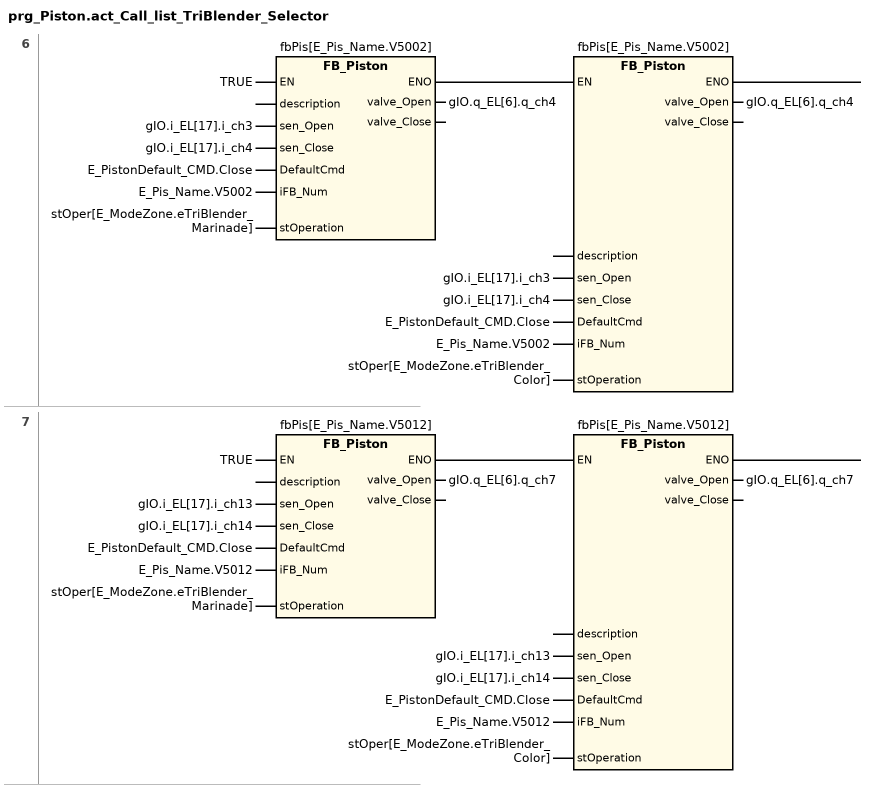
// NETWORK 6
fbPis[E_Pis_Name.V5002](
    sen_Open := gIO.i_EL[17].i_ch3,
    sen_Close := gIO.i_EL[17].i_ch4,
    DefaultCmd := E_PistonDefault_CMD.Close,
    iFB_Num := E_Pis_Name.V5002,
    stOperation := stOper[E_ModeZone.eTriBlender_Marinade],
    valve_Open => gIO.q_EL[6].q_ch4); // FB_Piston
fbPis[E_Pis_Name.V5002](
    sen_Open := gIO.i_EL[17].i_ch3,
    sen_Close := gIO.i_EL[17].i_ch4,
    DefaultCmd := E_PistonDefault_CMD.Close,
    iFB_Num := E_Pis_Name.V5002,
    stOperation := stOper[E_ModeZone.eTriBlender_Color],
    valve_Open => gIO.q_EL[6].q_ch4); // FB_Piston

// NETWORK 7
fbPis[E_Pis_Name.V5012](
    sen_Open := gIO.i_EL[17].i_ch13,
    sen_Close := gIO.i_EL[17].i_ch14,
    DefaultCmd := E_PistonDefault_CMD.Close,
    iFB_Num := E_Pis_Name.V5012,
    stOperation := stOper[E_ModeZone.eTriBlender_Marinade],
    valve_Open => gIO.q_EL[6].q_ch7); // FB_Piston
fbPis[E_Pis_Name.V5012](
    sen_Open := gIO.i_EL[17].i_ch13,
    sen_Close := gIO.i_EL[17].i_ch14,
    DefaultCmd := E_PistonDefault_CMD.Close,
    iFB_Num := E_Pis_Name.V5012,
    stOperation := stOper[E_ModeZone.eTriBlender_Color],
    valve_Open => gIO.q_EL[6].q_ch7); // FB_Piston
END_ACTION

ACTION act_Call_list_Water:
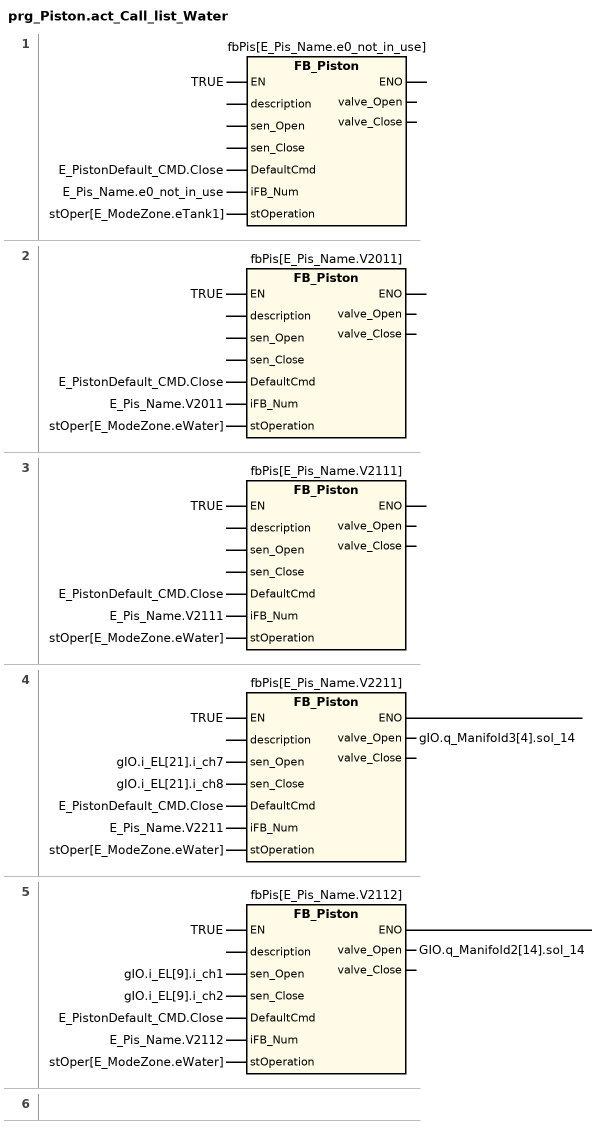
// NETWORK 1
fbPis[E_Pis_Name.e0_not_in_use](
    DefaultCmd := E_PistonDefault_CMD.Close,
    iFB_Num := E_Pis_Name.e0_not_in_use,
    stOperation := stOper[E_ModeZone.eTank1]); // FB_Piston

// NETWORK 2
fbPis[E_Pis_Name.V2011](
    DefaultCmd := E_PistonDefault_CMD.Close,
    iFB_Num := E_Pis_Name.V2011,
    stOperation := stOper[E_ModeZone.eWater]); // FB_Piston

// NETWORK 3
fbPis[E_Pis_Name.V2111](
    DefaultCmd := E_PistonDefault_CMD.Close,
    iFB_Num := E_Pis_Name.V2111,
    stOperation := stOper[E_ModeZone.eWater]); // FB_Piston

// NETWORK 4
fbPis[E_Pis_Name.V2211](
    sen_Open := gIO.i_EL[21].i_ch7,
    sen_Close := gIO.i_EL[21].i_ch8,
    DefaultCmd := E_PistonDefault_CMD.Close,
    iFB_Num := E_Pis_Name.V2211,
    stOperation := stOper[E_ModeZone.eWater],
    valve_Open => gIO.q_Manifold3[4].sol_14); // FB_Piston

// NETWORK 5
fbPis[E_Pis_Name.V2112](
    sen_Open := gIO.i_EL[9].i_ch1,
    sen_Close := gIO.i_EL[9].i_ch2,
    DefaultCmd := E_PistonDefault_CMD.Close,
    iFB_Num := E_Pis_Name.V2112,
    stOperation := stOper[E_ModeZone.eWater],
    valve_Open => GIO.q_Manifold2[14].sol_14); // FB_Piston

// NETWORK 6
END_ACTION

ACTION act_InterLock:
(*
IF TRUE 
AND stPis[E_Pis_Name.cheesy_cut].st_Deafult
AND stPis[E_Pis_Name.cheesy_down].st_Deafult
AND stPis[E_Pis_Name.cheesy_gripper].st_Deafult
AND stPis[E_Pis_Name.cheesy_turn].st_Deafult

AND stPis[E_Pis_Name.crown_down].st_Deafult
AND stPis[E_Pis_Name.crown_gripper].st_Deafult
AND stPis[E_Pis_Name.crown_press].st_Deafult
AND stPis[E_Pis_Name.crown_push].st_Deafult

AND stPis[E_Pis_Name.crust_down].st_Deafult
AND stPis[E_Pis_Name.crust_hold].st_Deafult
AND stPis[E_Pis_Name.crust_push].st_Deafult
AND stPis[E_Pis_Name.crust_roll].st_Deafult

AND stPis[E_Pis_Name.spikes_rotate_4].st_Deafult
AND stPis[E_Pis_Name.spikes_updown_4].st_Deafult

AND stPis[E_Pis_Name.door_4_2].st_Deafult

AND stPis[E_Pis_Name.trolley_down].st_Deafult

THEN;
	stPis[E_Pis_Name.trolley_move].b_InterLock:=TRUE;
ELSE;
	stPis[E_Pis_Name.trolley_move].b_InterLock:=FALSE;
END_IF
*)
END_ACTION

METHOD m_Disable_All : BOOL
VAR_INPUT
END_VAR

VAR
	i: INT;
END_VAR
FOR i:=1 TO E_Pis_Name.last DO;
	stPis[i].b_Enable:=FALSE;
END_FOR
END_METHOD

METHOD m_Enable_All : BOOL
VAR_INPUT
END_VAR

VAR
	i: INT;
END_VAR
FOR i:=1 TO E_Pis_Name.last DO;
	stPis[i].b_Enable:=TRUE;
END_FOR
END_METHOD

METHOD m_Get_Next_N : BOOL
VAR_IN_OUT
	iSel: INT;
END_VAR

VAR
	i: INT;
END_VAR

IF iSel> 1 THEN;
	FOR i:=iSel-1 TO 1 BY -1 DO
		IF stPis[i].b_Exist THEN;
			iSel:=i;
			RETURN;
		END_IF		
	END_FOR
END_IF
END_METHOD

METHOD m_Get_Next_P : BOOL
VAR_IN_OUT
	iSel: INT;
END_VAR

VAR
	i: INT;
END_VAR
//IF iSel< C_MAX_Pistons THEN;
//IF iSel< C_MAX_Pistons_Exist THEN;
IF iSel< E_Pis_Name.last THEN;
	FOR i:=iSel+1 TO E_Pis_Name.last BY 1 DO
		IF stPis[i].b_Exist THEN;
			iSel:=i;
			RETURN;
		END_IF		
	END_FOR
END_IF
END_METHOD

END_PROGRAM

// ---- 00 Library/01 Piston/FB_Piston.TcPOU
FUNCTION_BLOCK FB_Piston
VAR_INPUT
	description		: STRING;		(* Piston description*)	
	sen_Open		: BOOL;
	sen_Close		: BOOL;
	
	DefaultCmd		: E_PistonDefault_CMD:=E_PistonDefault_CMD.Close;

	iFB_Num			: E_Pis_Name;

END_VAR
VAR_OUTPUT
	valve_Open		: BOOL;
	valve_Close		: BOOL;	
END_VAR
VAR_IN_OUT
	stOperation		: ST_OperationButtons;	
END_VAR
VAR
	stPis			:	REFERENCE TO ST_Piston;
	stPis_UpLow		:	REFERENCE TO ST_Piston_U_L;
	state: E_Piston_State;
	state_Close,state_Open: (Ready, CheckState, ValveUpdate, Busy, Delay, Done, Error);

	//sen_Open_Exist	: REFERENCE TO BOOL :=FALSE;
	//sen_Close_Exist	: REFERENCE TO BOOL :=FALSE;
	
	ton_SensorCheck	: TON;
	ton_MinTime		: TON;
	ton_MaxTime		: TON;
	ton_SensorDelay	: TON;

	// Timing 
	t_minOpen		: TIME 	:=T#300MS;	(* minimum time to open piston*)
	t_minClose		: TIME	:=T#300MS;	(* minimum time to close piston*)
	t_maxOpen		: TIME 	:=T#3S;		(* Maximum time to open piston, will initiate an error*)
	t_maxClose		: TIME	:=T#3S;		(* Maximum time to open piston, will initiate an error*)
	t_DelayOpen		: TIME 	:=T#0S;		(* Delay time to getting "st_Open", will count after minimum time and sensors detection done*)
	t_DelayClose	: TIME	:=T#0S;		(* Delay time to getting "st_Close", will count after minimum time and sensors detection done*)	
	
	rt_Close		: R_TRIG;
	rt_Open			: R_TRIG;
	rt_OpenMan		: R_TRIG;
	rt_CloseMan		: R_TRIG;
	rt_DefaultPos	: R_TRIG;
	rt_ResumeMaster	: R_TRIG;
	b_memo_OpenFDBKExist	: BOOL;
	b_memo_CloseFDBKExist	: BOOL;
	Call_FTrig_ReqUp	: F_TRIG;
	Call_FTrig_ReqLow	: F_TRIG;
	
	bErrorMemo: BOOL;
		
	ton_Req_Close_timeout: TON;
	ton_Req_Open_timeout: TON;
	ton_Req_Default_timeout: TON;
	rt_StateSafe: R_TRIG;
	ft_StateSafe: F_TRIG;
END_VAR

IF iFB_Num <> E_Pis_Name.e0_not_in_use THEN;
	
END_IF

act_Get_Reference();




act_State_Machine();
act_StateDeafult();
//act_MemFdbkExist();

stPis_UpLow.bError:=stPis.b_Error;
stPis_UpLow.iFB_Num:=iFB_Num;
	
IF iFB_Num = E_Pis_Name.e0_not_in_use THEN;
	//stPis.st_Deafult:=TRUE;
END_IF


rt_StateSafe(CLK:=stOperation.bStateSafe_mode);
ft_StateSafe(CLK:=stOperation.bStateSafe_mode);

IF __ISVALIDREF(stPis) THEN;
	IF ft_StateSafe.Q
	AND NOT stPis.st_Deafult
	THEN;
		//stPis.req_DefaultPos:=TRUE;
		//stPis.req_Close:=FALSE;
		//stPis.req_Open:=FALSE;	
	END_IF
	
	IF rt_StateSafe.Q THEN;
		
		IF NOT stPis.st_Deafult THEN;
			//stPis.req_DefaultPos:=TRUE;
		END_IF	
		stPis.b_Resume:=TRUE;
		//stPis.b_Reset:=TRUE;	
	END_IF	
END_IF

ACTION act_Close:



CASE state_Close OF
	Ready:;
		IF stPis.req_CloseMan THEN;
			stPis.req_CloseMan:=FALSE;
			// Do manual case code
			stPis.req_Close:=TRUE;
		END_IF		
		IF stPis.req_Close THEN;
			stPis.req_Open:=FALSE;
			stPis.req_OpenMan:=FALSE;	
			stPis.req_DefaultPos:=FALSE;			
			state_Close:=CheckState;
		END_IF
		
	CheckState:;
		IF stPis.st_Close THEN;
			stPis.st_Open:=FALSE;
			state_Close:=Done;
		ELSE;
			stPis.st_Close:=FALSE;
			stPis.st_Open:=FALSE;
			state_Close:=ValveUpdate;
		END_IF
		
	ValveUpdate:;
		valve_Open:=FALSE;
		valve_Close:=TRUE;
		ton_SensorCheck(IN:=FALSE);
		ton_MinTime(IN:=FALSE);
		ton_MinTime(IN:=TRUE);
		ton_MaxTime(IN:=FALSE);
		ton_MaxTime(IN:=TRUE);
		ton_SensorDelay(IN:=FALSE);
		
		stPis.t_LastClose:=T#0S;
		state_Close:=Busy;
		
	Busy:;
		ton_MinTime(PT:=t_minClose);
		ton_MaxTime(PT:=t_maxClose, IN:=TRUE);
		ton_SensorDelay(PT:=t_DelayClose,IN:=m_PistonSensorCheck());	
		IF 	ton_MinTime.Q 		
		AND ton_SensorDelay.IN THEN;
			ton_MaxTime(IN:=FALSE);
			IF ton_SensorDelay.Q THEN;
				stPis.t_LastClose:=ton_MaxTime.ET;			
				state_Close:=Done;				
			END_IF
		ELSE;
			IF ton_MaxTime.Q THEN;
				//Error to print
				state_Close:=Error;
			END_IF			
		END_IF
	
	Done:;
		stPis.st_Close:=TRUE;
		IF stPis.st_Close THEN;
			state_Close:=Ready;
			stPis.req_Close:=FALSE;
		END_IF	
		
	Error:;
		//Wating to operator reset & resume 
		stPis.b_Error:=TRUE;	
		m_Error();
		IF stPis.b_Resume THEN;
			state_Close:=ValveUpdate;
			//stPis.b_Resume:=FALSE;	
			//stPis.b_Error:=FALSE;
			//bErrorMemo:=FALSE;
		END_IF
		
END_CASE
END_ACTION

ACTION act_Get_Reference:
stPis REF= g_Piston.stPis[iFB_Num];
stPis_UpLow REF= g_Piston.stPis_U_L[iFB_Num];
//stPis.description:=description;
stPis.b_Exist:=TRUE;
stPis.sName:=TO_STRING(iFB_Num);
stPis.iPisNum:=iFB_Num;
arPisName[iFB_Num].Num:=iFB_Num;
arPisName[iFB_Num].Description:=stPis.sName;

stPis.sen_Close REF= sen_Close;
stPis.sen_Close_Exist REF= stPisSetting[iFB_Num].sen_Close_Exist;
//stPis.sen_Close_Exist REF= sen_Close_Exist;
stPis.sen_Open REF= sen_Open;
stPis.sen_Open_Exist REF= stPisSetting[iFB_Num].sen_Open_Exist;
//stPis.sen_Open_Exist REF= sen_Open_Exist;

stPis.valve_Close REF= valve_Close;
stPis.valve_Open REF= valve_Open;

stPis.t_maxClose REF= stPisSetting[iFB_Num].t_maxClose;
stPis.t_maxOpen REF= stPisSetting[iFB_Num].t_maxOpen;
stPis.t_minClose REF= stPisSetting[iFB_Num].t_minClose;
stPis.t_minOpen REF= stPisSetting[iFB_Num].t_minOpen;
stPis.t_DelayClose REF= stPisSetting[iFB_Num].t_DelayClose;
stPis.t_DelayOpen REF= stPisSetting[iFB_Num].t_DelayOpen;
t_maxClose:=fun_Real_SecondsToTime(in_Time:=stPis.t_maxClose);
t_maxOpen:=fun_Real_SecondsToTime(in_Time:=stPis.t_maxOpen);
t_minClose:=fun_Real_SecondsToTime(in_Time:=stPis.t_minClose);
t_minOpen:=fun_Real_SecondsToTime(in_Time:=stPis.t_minOpen);
t_DelayClose:=fun_Real_SecondsToTime(in_Time:=stPis.t_DelayClose);
t_DelayOpen:=fun_Real_SecondsToTime(in_Time:=stPis.t_DelayOpen);

stPis.DefaultCmd REF= DefaultCmd;

IF stPis.b_Error THEN;
	stOperation.bSetPause:=TRUE;
END_IF
(*
IF stPis.b_Error 
AND stDevErr_H.eErrorActive=E_Error_Active_Module.noError 
THEN;
	stDevErr_H.sObjectName:=CONCAT('pis.No:',INT_TO_STRING(stPis.iPisNum));
	stDevErr_H.sObjectName:=CONCAT(stDevErr_H.sObjectName,'- ');
	stDevErr_H.sObjectName:=CONCAT(stDevErr_H.sObjectName,TO_STRING(iFB_Num));
	stDevErr_H.eErrorActive:=E_Error_Active_Module.Piston;
	stDevErr_H.iObjectID:=iFB_Num;
END_IF

rt_ResumeMaster(CLK:=stDevErr_H.bMasterResume);
IF rt_ResumeMaster.Q THEN;
	stPis.b_Resume:=TRUE;
END_IF
*)
END_ACTION

ACTION act_MemFdbkExist:
IF stPis.valve_Close AND stPis_UpLow.exist THEN
	//Fetching signals
	IF TRUE THEN
		Call_FTrig_ReqUp(CLK:=stPis_UpLow.req_Upper , Q=> );
	ELSE
		Call_FTrig_ReqUp(CLK:=stPis_UpLow.st_Upper , Q=> );
	END_IF
	
	Call_FTrig_ReqLow(CLK:=stPis_UpLow.st_Lower , Q=> );
	
	//setting memmory
	IF stPis_UpLow.req_Lower AND stPis.sen_Close_Exist THEN
		b_memo_CloseFDBKExist:=stPis.sen_Close_Exist;
		stPis.sen_Close_Exist:=FALSE;
	ELSIF stPis_UpLow.req_Lower AND b_memo_CloseFDBKExist THEN
		stPis.sen_Close_Exist:=FALSE;
	END_IF
	
	IF stPis_UpLow.req_Upper AND stPis.sen_Open_Exist THEN
		b_memo_OpenFDBKExist:=stPis.sen_Open_Exist;
		stPis.sen_Open_Exist:=FALSE;
	ELSIF stPis_UpLow.req_Upper AND b_memo_OpenFDBKExist THEN
		stPis.sen_Open_Exist:=FALSE;
	END_IF
	//resseting memmory
	IF Call_FTrig_ReqUp.Q AND b_memo_OpenFDBKExist THEN
		stPis.sen_Open_Exist:=b_memo_OpenFDBKExist;
		b_memo_OpenFDBKExist:=FALSE;
	END_IF
	
	IF Call_FTrig_ReqLow.Q AND b_memo_CloseFDBKExist THEN
		stPis.sen_Close_Exist:=b_memo_CloseFDBKExist;
		b_memo_CloseFDBKExist:=FALSE;
	END_IF
ELSE
	IF stPis_UpLow.exist THEN
		b_memo_CloseFDBKExist:=FALSE;
		b_memo_OpenFDBKExist:=FALSE;
		stPis_UpLow.req_Lower:=FALSE;
		stPis_UpLow.st_Lower:=FALSE;
	ELSE
		;
	END_IF
	
END_IF

IF stPis.req_Open AND NOT stPis_UpLow.exist  THEN
	IF stPis.sen_Close_Exist THEN
		b_memo_CloseFDBKExist:=TRUE;
		stPis.sen_Close_Exist:=FALSE;
	END_IF
	
	IF stPis.sen_Open_Exist THEN
		b_memo_OpenFDBKExist:=TRUE;
		stPis.sen_Open_Exist:=FALSE;
	END_IF
ELSIF stPis.req_Close AND NOT stPis_UpLow.exist THEN
	IF b_memo_CloseFDBKExist THEN
		stPis.sen_Close_Exist:=TRUE;
		b_memo_CloseFDBKExist:=FALSE;
	END_IF
	
	IF b_memo_OpenFDBKExist THEN
		stPis.sen_Open_Exist:=TRUE;
		b_memo_OpenFDBKExist:=FALSE;
	END_IF
	
END_IF
END_ACTION

ACTION act_New_CMD:
IF stPis.b_Enable AND stPis.b_InterLock THEN;
	
	rt_Close(CLK:=stPis.req_Close AND NOT ton_Req_Close_timeout.Q);
	rt_Open(CLK:=stPis.req_Open AND NOT ton_Req_Open_timeout.Q);
	rt_CloseMan(CLK:=stPis.req_CloseMan);
	rt_OpenMan(CLK:=stPis.req_OpenMan);
	rt_DefaultPos(CLK:=stPis.req_DefaultPos AND NOT ton_Req_Default_timeout.Q);
	
	ton_Req_Close_timeout(PT:=T#0.1S);	
	IF (stPis.req_Close OR stPis.req_CloseMan)
	AND state_Close=Ready
	AND NOT ton_Req_Close_timeout.Q
	THEN;
		ton_Req_Close_timeout.IN:=TRUE;
	ELSE;
		ton_Req_Close_timeout.IN:=FALSE;
	END_IF

	ton_Req_Open_timeout(PT:=T#0.1S);	
	IF (stPis.req_Open OR stPis.req_OpenMan)
	AND state_Open=Ready
	AND NOT ton_Req_Open_timeout.Q
	THEN;
		ton_Req_Open_timeout.IN:=TRUE;
	ELSE;
		ton_Req_Open_timeout.IN:=FALSE;
	END_IF

	ton_Req_Default_timeout(PT:=T#0.1S);	
	IF (stPis.req_DefaultPos OR stPis.req_DefaultPos)
	AND state_Open=Ready
	AND NOT ton_Req_Default_timeout.Q
	THEN;
		ton_Req_Default_timeout.IN:=TRUE;
	ELSE;
		ton_Req_Default_timeout.IN:=FALSE;
	END_IF
	
	IF rt_Close.Q OR rt_CloseMan.Q THEN; 
		state:=E_Piston_State.Busy_Close; 
		stPis.req_Open:=FALSE;
		stPis.req_OpenMan:=FALSE;	
		stPis.req_DefaultPos:=FALSE;	
	END_IF
	IF rt_Open.Q OR rt_OpenMan.Q THEN; 
		state:=E_Piston_State.Busy_Open; 
		stPis.req_Close:=FALSE;
		stPis.req_CloseMan:=FALSE;
		stPis.req_DefaultPos:=FALSE;	
	END_IF
	IF rt_DefaultPos.Q THEN; 
		state:=E_Piston_State.Init; 
	END_IF
	
	(*IF rt_CloseMan.Q THEN; 
		state:=E_Piston_State.Busy_Close;
	END_IF
	IF rt_OpenMan.Q THEN; 
		state:=E_Piston_State.Busy_Open; 
	END_IF
*)
	
	IF rt_Close.Q 
	OR rt_Open.Q
	OR rt_CloseMan.Q
	OR rt_OpenMan.Q
	OR rt_DefaultPos.Q
	THEN;
		stPis.b_Error:=FALSE;
		bErrorMemo:=FALSE;
	END_IF
	
	stPis.b_DeactivateMan:=FALSE;
ELSE;
	stPis.b_DeactivateMan:=TRUE;
END_IF
END_ACTION

ACTION act_Open:



CASE state_Open OF
	Ready:;
		IF stPis.req_OpenMan THEN;
			stPis.req_OpenMan:=FALSE;
			// Do manual case code
			stPis.req_Open:=TRUE;
		END_IF		
		IF stPis.req_Open THEN;
			stPis.req_Close:=FALSE;
			stPis.req_CloseMan:=FALSE;
			stPis.req_DefaultPos:=FALSE;		
			state_Open:=CheckState;
		END_IF
		
	CheckState:;
		IF stPis.st_Open THEN;
			stPis.st_Close:=FALSE;
			state_Open:=Done;
		ELSE;
			stPis.st_Close:=FALSE;
			stPis.st_Open:=FALSE;
			state_Open:=ValveUpdate;
		END_IF
		
	ValveUpdate:;
		valve_Open:=TRUE;
		valve_Close:=FALSE;
		ton_SensorCheck(IN:=FALSE);
		ton_MinTime(IN:=FALSE);
		ton_MinTime(IN:=TRUE);
		ton_MaxTime(IN:=FALSE);
		ton_MaxTime(IN:=TRUE);	
		ton_SensorDelay(IN:=FALSE);
		
		stPis.t_LastOpen:=T#0S;	
		state_Open:=Busy;
		
	Busy:;
		ton_MinTime(PT:=t_minOpen);
		ton_MaxTime(PT:=t_maxOpen);
		ton_SensorDelay(PT:=t_DelayOpen,IN:=m_PistonSensorCheck());	
		IF 	ton_MinTime.Q 
		AND m_PistonSensorCheck()	THEN;
			ton_MaxTime(IN:=FALSE);
			IF ton_SensorDelay.Q THEN;
				stPis.t_LastOpen:=ton_MaxTime.ET;			
				state_Open:=Done;				
			END_IF
		ELSE;
			IF ton_MaxTime.Q THEN;
				//Error to print
				state_Open:=Error;
				;
			END_IF				
		END_IF
	
	Done:;
		stPis.st_Open:=TRUE;	
		IF stPis.st_Open THEN;
			state_Open:=Ready;
			stPis.req_Open:=FALSE;
		END_IF	
		
	Error:;
		//Wating to operator reset & resume 
		stPis.b_Error:=TRUE;
		m_Error();
		IF stPis.b_Resume THEN;
			state_Open:=ValveUpdate;
			//stPis.b_Resume:=FALSE;
			//stPis.b_Error:=FALSE;
			//bErrorMemo:=FALSE;
		END_IF
		
END_CASE
END_ACTION

ACTION act_State_Machine:
IF stPis.b_Resume THEN;
	stPis.b_Error:=FALSE;
	bErrorMemo:=FALSE;		
END_IF

act_New_CMD();
CASE state OF
	E_Piston_State.Init:;
			ton_SensorCheck(IN:=FALSE);
			
	
			stPis.st_Close:=FALSE;
			stPis.st_Open:=FALSE;
			
			stPis.b_Error:=FALSE;
			stPis.b_Reset:=FALSE;
			stPis.b_Resume:=FALSE;
			
			stPis.req_Close:=FALSE;
			stPis.req_CloseMan:=FALSE;	
			stPis.req_Open:=FALSE;
			stPis.req_OpenMan:=FALSE;
			stPis.req_DefaultPos:=FALSE;
			
			state_Close:=Ready;
			state_Open:=Ready;
			
			//check default configuration
			IF stPis.b_Enable AND stPis.b_InterLock THEN;				
				CASE DefaultCmd OF
					E_PistonDefault_CMD.Close:;
						state:=E_Piston_State.Busy_Close;
						stPis.req_Close:=TRUE;
					E_PistonDefault_CMD.Open:;
						state:=E_Piston_State.Busy_Open;
						stPis.req_Open:=TRUE;
					E_PistonDefault_CMD.Sensors:;
					E_PistonDefault_CMD.SensorsClose:;
					E_PistonDefault_CMD.SensorsOpen:;
					
				END_CASE
			END_IF
	
	E_Piston_State.Close:;
		IF m_PistonSensorCheck() AND NOT stPis.b_Error THEN;
			stPis.st_Close:=TRUE;
			stPis.st_Open:=FALSE;
			ton_SensorCheck(IN:=FALSE);
		ELSE;
			ton_SensorCheck(IN:=TRUE);
			IF ton_SensorCheck.Q THEN;
				stPis.st_Close:=FALSE;
				stPis.st_Open:=FALSE;				
				stPis.b_Error:=TRUE;
				m_Error();		
			END_IF			
		END_IF
				
	E_Piston_State.Open:;
		IF m_PistonSensorCheck() AND NOT stPis.b_Error THEN;
			stPis.st_Close:=FALSE;
			stPis.st_Open:=TRUE;
			ton_SensorCheck(IN:=FALSE);
		ELSE;			
			ton_SensorCheck(IN:=TRUE);
			IF ton_SensorCheck.Q THEN;
				stPis.st_Close:=FALSE;
				stPis.st_Open:=FALSE;				
				stPis.b_Error:=TRUE;
				m_Error();
			END_IF
		END_IF
	
	E_Piston_State.Busy_Close:;
		ton_SensorCheck(IN:=FALSE);
		act_Close();		
		state_Open:=Ready;		
		IF stPis.st_Close AND NOT stPis.req_Close THEN;
			state:=E_Piston_State.Close;
		END_IF

	E_Piston_State.Busy_Open:;
		ton_SensorCheck(IN:=FALSE);
		act_Open();
		state_Close:=Ready;
		IF stPis.st_Open AND NOT stPis.req_Open THEN;
			state:=E_Piston_State.Open;
		END_IF
END_CASE			

ton_SensorCheck(PT:=T#4S);//PT:=T#0.5S

IF ton_SensorCheck.Q THEN;
	stPis.b_Error:=TRUE;		
END_IF
stPis.b_Resume:=FALSE;
END_ACTION

ACTION act_StateDeafult:
CASE DefaultCmd	OF
	E_PistonDefault_CMD.Close:;
		stPis.st_Deafult:=stPis.st_Close;
	E_PistonDefault_CMD.Open:;
		stPis.st_Deafult:=stPis.st_Open;
END_CASE
END_ACTION

METHOD PUBLIC m_CheckByRecipe : BOOL
VAR_INPUT
	stPis: ST_Piston;
	req: E_Piston_Recipe_State;	
END_VAR
m_CheckByRecipe:=FALSE;
IF stPis.iPisNum <> E_Pis_Name.e0_not_in_use THEN
	CASE req OF
		E_Piston_Recipe_State.NoChanges:;
			m_CheckByRecipe:=TRUE;
		E_Piston_Recipe_State.Act:;
			IF (stPis.DefaultCmd=E_PistonDefault_CMD.Close AND stPis.st_Open) 
			OR (stPis.DefaultCmd=E_PistonDefault_CMD.Open AND stPis.st_Close)
			THEN;
				m_CheckByRecipe:=TRUE;
			END_IF
		E_Piston_Recipe_State.Release:;
			IF (stPis.DefaultCmd=E_PistonDefault_CMD.Close AND stPis.st_Close) 
			OR (stPis.DefaultCmd=E_PistonDefault_CMD.Open AND stPis.st_Open)
			THEN;
				m_CheckByRecipe:=TRUE;
			END_IF	
	END_CASE
ELSE;
	m_CheckByRecipe:=TRUE;
END_IF
END_METHOD

METHOD m_Error : BOOL
VAR_INPUT
END_VAR
VAR
	sActErrorID_AA: STRING;
	sActErrorID: STRING;
	Mess: INT;
	cFound: INT;
	iFound: INT;
	i: INT;
	bWarning: BOOL;

END_VAR
(*
IF SFCError OR bWarning THEN

	IF  SFCErrorStep='WaitSenOpen' THEN
		stPis.eErrNum:=1;
	ELSIF SFCErrorStep='WaitSenNotClose' THEN
		stPis.eErrNum:=2;
	ELSIF SFCErrorStep='WaitSenClose' THEN
		stPis.eErrNum:=3;
	ELSIF SFCErrorStep='WaitSenNotOpen' THEN
		stPis.eErrNum:=4;
	ELSIF SFCErrorStep='No Status' THEN
		stPis.eErrNum:=5;
	ELSIF SFCErrorStep='No Valve Operation' THEN
		stPis.eErrNum:=6;
	ELSIF SFCErrorStep='Not synchronized with cycle command' THEN //SensorsChecking
		stPis.eErrNum:=7;
	ELSIF SFCErrorStep='SensorsChecking' THEN
		stPis.eErrNum:=8;		
	ELSIF bWarning THEN;	// act_Ready
		//stPis.eErrNum:=21; 	// '2AAx021',	'Warning',	', Manual command rejected in semi/auto mode',	(**)
	ELSE
		stPis.eErrNum:=9;
	END_IF
	Last_SFCErrorStep:=SFCErrorStep;
	
ELSE
		stPis.eErrNum:=0;
END_IF
*)
// Temp solution
IF stPis.b_Error THEN;
	stPis.eErrNum:=1;
END_IF

IF stPis.eErrNum<>0 AND NOT bErrorMemo AND stPis.iPisNum<>0 THEN

	IF stPis.iPisNum<10 THEN
		sActErrorID:=CONCAT('20',INT_TO_STRING(stPis.iPisNum));
	ELSE
		sActErrorID:=CONCAT('2',INT_TO_STRING(stPis.iPisNum));
	END_IF
	
	IF stPis.eErrNum<10 THEN
		sActErrorID:=CONCAT(sActErrorID,'x00');
		sActErrorID:=CONCAT(sActErrorID,INT_TO_STRING(stPis.eErrNum));
	ELSE
		sActErrorID:=CONCAT(sActErrorID,'x0');
		sActErrorID:=CONCAT(sActErrorID,INT_TO_STRING(stPis.eErrNum));		
	END_IF

	FOR Mess:=100 TO 2 BY -1 DO
		Buffer_Act_Message[Mess].sDateTime:=Buffer_Act_Message[Mess-1].sDateTime;
		Buffer_Act_Message[Mess].sErrID:=Buffer_Act_Message[Mess-1].sErrID;
		Buffer_Act_Message[Mess].sLevel:=Buffer_Act_Message[Mess-1].sLevel;
		Buffer_Act_Message[Mess].sModuleDescription:=Buffer_Act_Message[Mess-1].sModuleDescription;
		Buffer_Act_Message[Mess].sErrorMessage:=Buffer_Act_Message[Mess-1].sErrorMessage;
	END_FOR
		Buffer_Act_Message[1].sDateTime:=sRealTime;
		Buffer_Act_Message[1].sErrID:=sActErrorID;
		Buffer_Act_Message[1].sLevel:='Error';
		//Buffer_Act_Message[1].sModuleDescription:='Pneumatic valve';
		Buffer_Act_Message[1].sModuleDescription:=stOperation.sModeZone;

		(*888888888888888888888888888888888888888888*)
		IF stPis.eErrNum<10 THEN
			sActErrorID_AA:=CONCAT('2AAx00',INT_TO_STRING(stPis.eErrNum));
		ELSE
			sActErrorID_AA:=CONCAT('2AAx0',INT_TO_STRING(stPis.eErrNum));			
		END_IF
		cFound:=0;
		FOR i:=1 TO C_Max_ErrorList DO
			IF ar_ErrorList[i,eErrID]=sActErrorID_AA THEN
				iFound:=i;
				ar_ErrorActive[iFound]:=TRUE;
				cFound:=cFound+1;
			END_IF
		END_FOR

		Buffer_Act_Message[1].sErrorMessage:=CONCAT( 'Piston Num ', INT_TO_STRING(stPis.iPisNum));
		Buffer_Act_Message[1].sErrorMessage:=CONCAT( Buffer_Act_Message[1].sErrorMessage, ', ');
		//Buffer_Act_Message[1].sErrorMessage:=CONCAT( Buffer_Act_Message[1].sErrorMessage, arPisDescription[stPis.iPisNum]);
		Buffer_Act_Message[1].sErrorMessage:=CONCAT( Buffer_Act_Message[1].sErrorMessage, stPis.sName);
		Buffer_Act_Message[1].sErrorMessage:=CONCAT( Buffer_Act_Message[1].sErrorMessage, ': ');

		IF cFound=1 THEN;
			Buffer_Act_Message[1].sErrorMessage:=CONCAT( Buffer_Act_Message[1].sErrorMessage, ar_ErrorList[iFound,eErrMeassage]);	(*	Error from the List	*)
			Buffer_Act_Message[1].sLevel:= ar_ErrorList[iFound,eErrLevel];	(*	Level from the List	*)
		ELSIF cFound=0 THEN;
			Buffer_Act_Message[1].sErrorMessage:=CONCAT( Buffer_Act_Message[1].sErrorMessage, 'Error ID not found on the "Error_List"');	(*	Error ID not Foud on the List	*)
		ELSIF cFound>1 THEN;
			Buffer_Act_Message[1].sErrorMessage:=CONCAT( Buffer_Act_Message[1].sErrorMessage, 'More then one error with the same ID  found on the "Error_list"');	(*	More then one Errors Foud with the same  ID		*)
		END_IF
		(*888888888888888888888888888888888888888888*)

	FUN_Write_Line_To_History();
	bErrorMemo:=TRUE;
END_IF

(*
'WaitSenOpen'
'WaitSenNotClose'
'WaitSenClose'
'WaitSenNotOpen'
'No Status'
'No Valve Operation'
*)
END_METHOD

METHOD m_PistonSensorCheck : BOOL
(*VAR_INPUT
	exist: BOOL;
	SensorState: BOOL;
	ValveState: BOOL;

END_VAR*)
VAR
	OK_Open: BOOL;
	OK_Close: BOOL;


END_VAR
IF stPis.sen_Close_Exist THEN;

	//IF valve_Close = sen_Close THEN;
	IF valve_Close THEN;
		IF stPis_UpLow.out_Upper OR stPis_UpLow.out_Lower THEN;
			OK_Close:=TRUE;
		ELSE;
			OK_Close:=sen_Close;
		END_IF
	ELSE ;
		OK_Close:=NOT sen_Close;
	END_IF
ELSE
	OK_Close:=TRUE;
END_IF

IF stPis.sen_Open_Exist THEN;
	IF valve_Open = sen_Open THEN;
		OK_Open:=TRUE;	
	ELSE;
		OK_Open:=FALSE;
	END_IF
ELSE
	OK_Open:=TRUE;
END_IF

IF OK_Close AND OK_Open THEN;
	m_PistonSensorCheck:=TRUE;
ELSE;
	m_PistonSensorCheck:=FALSE;
END_IF
END_METHOD

METHOD PUBLIC m_SetByRecipe : BOOL
VAR_INPUT
	
	req: E_Piston_Recipe_State;
END_VAR
VAR
	ref_stPis: REFERENCE TO ST_Piston;
END_VAR

VAR_IN_OUT
	stPis: ST_Piston;
END_VAR
IF stPis.iPisNum <> E_Pis_Name.e0_not_in_use THEN
	//ref_stPis REF= stPis;
	CASE req OF
		E_Piston_Recipe_State.NoChanges:;
			//Done
		E_Piston_Recipe_State.Act:;
			IF stPis.DefaultCmd=E_PistonDefault_CMD.Close THEN;
				IF NOT stPis.st_Open THEN;
					stPis.req_Open:=TRUE;
				END_IF		
			ELSIF stPis.DefaultCmd=E_PistonDefault_CMD.Open THEN;
				IF NOT stPis.st_Close THEN;
					stPis.req_Close:=TRUE;
				END_IF				
			END_IF
	
		E_Piston_Recipe_State.Release:;
			IF stPis.DefaultCmd=E_PistonDefault_CMD.Close THEN;
				IF NOT stPis.st_Close THEN;
					stPis.req_Close:=TRUE;
				END_IF			
			ELSIF stPis.DefaultCmd=E_PistonDefault_CMD.Open THEN;
				IF NOT stPis.st_Open THEN;
					stPis.req_Open:=TRUE;
				END_IF			
			END_IF	
	END_CASE	
END_IF
END_METHOD

END_FUNCTION_BLOCK

// ---- 00 Library/10 Utils/fun_Real_SecondsToTime.TcPOU
FUNCTION fun_Real_SecondsToTime : TIME
VAR_INPUT
	in_Time: REAL; // Seconds

END_VAR
VAR
END_VAR

fun_Real_SecondsToTime:=DINT_TO_TIME(TRUNC(in_Time*1000));

END_FUNCTION

// ---- 00 Library/04-Messages/FUN_Write_Line_To_History.TcPOU
FUNCTION FUN_Write_Line_To_History : BOOL
VAR_INPUT
END_VAR
VAR
	i: INT;
END_VAR

	FOR i:=C_Max_Buffer_Act_list TO 2 BY -1 DO
		Buffer_Act_History[i]:=Buffer_Act_History[i-1];
	END_FOR
	Buffer_Act_History[1]:=Buffer_Act_Message[1];

END_FUNCTION

// ---- 00 Library/01 Piston/FB_Piston_U_L.TcPOU
FUNCTION_BLOCK PUBLIC FB_Piston_U_L// EXTENDS FB_Piston
VAR_INPUT
	enable		: BOOL	;
	sen_Upper	: BOOL	;
	sen_Lower	: BOOL	;

END_VAR
VAR_OUTPUT
	valve_Upper		:BOOL;
	valve_Lower		:BOOL;	
END_VAR
VAR
	tOn: TIME:=T#1S;
	tOff: TIME:=T#1S;
	Call_RTrig_ReqUp: R_TRIG;
	Call_RTrig_ReqLow: R_TRIG;
	
	b_Memo_ReqUp	:	BOOL	;
	b_Memo_ReqLow	:	BOOL	;
	Call_FTrig_Error: 	F_TRIG	;
	stPis			:	REFERENCE TO ST_Piston;
	ton_req_Upper: TON;
	ton_req_Lower: TON;
	tOperation: TIME := T#2S;
	ton_err_Upper: TON;
	ton_err_Lower: TON;
	tError: TIME := T#5s;
END_VAR
VAR_IN_OUT
	st_Piston_U_L	:	ST_Piston_U_L	;
	stOperation		: ST_OperationButtons;
END_VAR

act_Get_Reference();
act_SetOutputs();

IF stPis.b_Error THEN;
	stOperation.bSetPause:=TRUE;
END_IF

ton_req_Upper(PT:=tOperation, IN:=st_Piston_U_L.req_Upper);
ton_req_Lower(PT:=tOperation, IN:=st_Piston_U_L.req_Lower);

ton_err_Upper(PT:=tError);
ton_err_Lower(PT:=tError);

IF TRUE 
AND st_Piston_U_L.req_Upper
AND (NOT st_Piston_U_L.st_Upper)
AND (NOT FALSE) // reset error
THEN;
	ton_err_Upper.IN:=TRUE;
ELSE;
	ton_err_Upper.IN:=FALSE;
END_IF

IF TRUE 
AND st_Piston_U_L.req_Lower
AND (NOT st_Piston_U_L.st_Lower)
AND (NOT FALSE) // reset error
THEN;
	ton_err_Lower.IN:=TRUE;
ELSE;
	ton_err_Lower.IN:=FALSE;
END_IF

IF ton_err_Upper.Q OR ton_err_Lower.Q THEN;
	stPis.b_Error:=TRUE;
END_IF

ACTION act_Get_Reference:
//st_Piston_U_L.str_Piston REF= g_Piston.stPis[iFB_Num];
stPis REF= g_Piston.stPis[st_Piston_U_L.iFB_Num];
END_ACTION

ACTION act_SetOutputs:
(*IF st_Piston_U_L.bError THEN
	IF st_Piston_U_L.req_Upper THEN
		b_Memo_ReqUp:=TRUE;
	END_IF
	IF st_Piston_U_L.req_Lower THEN
		b_Memo_ReqLow:=TRUE;
	END_IF
	st_Piston_U_L.req_Upper:=FALSE;
	st_Piston_U_L.req_Lower:=FALSE;
END_IF*)

(*
Call_FTrig_Error(CLK:=st_Piston_U_L.bError , Q=> );

IF Call_FTrig_Error.Q THEN
	st_Piston_U_L.req_Upper:=b_Memo_ReqUp;
	st_Piston_U_L.req_Lower:=b_Memo_ReqLow;
	b_Memo_ReqUp:=FALSE;
	b_Memo_ReqLow:=FALSE;
END_IF*)

//Resseting opposite signal
//***************************************************************
Call_RTrig_ReqUp(CLK:=st_Piston_U_L.req_Upper , Q=> );
Call_RTrig_ReqLow(CLK:=st_Piston_U_L.req_Lower, Q=> );
IF Call_RTrig_ReqUp.Q THEN
	st_Piston_U_L.req_Lower:=FALSE;
END_IF

IF Call_RTrig_ReqLow.Q THEN
	st_Piston_U_L.req_Upper :=FALSE;
END_IF
//***************************************************************

IF enable AND stPis.valve_Close THEN;
	st_Piston_U_L.exist:=TRUE;
	
	IF st_Piston_U_L.req_Upper THEN;
		valve_Upper:=TRUE;
		valve_Lower:=FALSE;		
	ELSIF st_Piston_U_L.req_Lower THEN;
		valve_Upper:=FALSE;
		valve_Lower:=TRUE;		
	ELSE;
		valve_Upper:=FALSE;
		valve_Lower:=FALSE;		
	END_IF
ELSE;
	st_Piston_U_L.exist:=FALSE;
	st_Piston_U_L.req_Upper:=FALSE;
	st_Piston_U_L.req_Lower:=FALSE;
	valve_Upper:=FALSE;
	valve_Lower:=FALSE;
END_IF

//outputs for hmi
st_Piston_U_L.out_Upper:=valve_Upper;
st_Piston_U_L.out_Lower:=valve_Lower;

//Status
st_Piston_U_L.st_Upper:=m_sen_Upper();
st_Piston_U_L.st_Lower:=m_sen_Lower();
st_Piston_U_L.st_Released:=(NOT m_sen_Upper() AND NOT m_sen_Lower());

st_Piston_U_L.sen_Upper:=sen_Upper;
st_Piston_U_L.sen_Lower:=sen_Lower;
END_ACTION

METHOD m_sen_Lower : BOOL
VAR_INPUT
END_VAR
IF st_Piston_U_L.sen_Lower_exist THEN; // sensor exist
	m_sen_Lower:=sen_Lower;
ELSE;
	m_sen_Lower:=ton_req_Lower.Q;
END_IF
END_METHOD

METHOD m_sen_Upper : BOOL
VAR_INPUT
END_VAR
IF st_Piston_U_L.sen_Upper_exist THEN; // sensor exist
	m_sen_Upper:=sen_Upper;
ELSE;
	m_sen_Upper:=ton_req_Upper.Q;
END_IF
END_METHOD

END_FUNCTION_BLOCK

// ---- 00 Library/05 Safety/prg_Safety.TcPOU
PROGRAM prg_Safety
VAR
	(*
	rt_TSafe_OK: R_TRIG;
	rt_TSafe_Err: R_TRIG;
	ton_TSafe_OK: TON;
	ton_TSafe_Err_Reset_ON: TON;
	ton_TSafe_Err_Reset_OFF: TON;
	*)
	fbTwinSAFE: ARRAY[1..1] OF FB_TwinSAFE;
	
	HMI_ES1_Restart: BOOL;
	HMI_ES2_Restart: BOOL;
	HMI_ES3_Restart: BOOL;
	HMI_ES4_Restart: BOOL;
	
	rtStateSafe: R_TRIG;
	ftStateSafe: F_TRIG;
END_VAR


act_Call_TSs();


{IF defined (Production)}
	bStateSafe_ES1:=arSafe[1].stSafetyIn.ES1_State;
	//bStateSafe_ES2:=arSafe[1].stSafetyIn.ES2_State;
	bStateSafe_ES3:=arSafe[1].stSafetyIn.ES3_State;
	//bStateSafe_ES4:=arSafe[1].stSafetyIn.ES4_State;
{ELSIF defined (Simulation_IO)}
	bES_Bypass:= TRUE;

	bStateSafe_ES1:=TRUE;
	bStateSafe_ES2:=TRUE;
	bStateSafe_ES3:=TRUE;
	bStateSafe_ES4:=TRUE;
{END_IF}

IF TRUE 
AND bStateSafe_ES1
//AND bStateSafe_ES2
AND bStateSafe_ES3
//AND bStateSafe_ES4

OR bES_Bypass

THEN;
	bStateSafe:=TRUE;
ELSE;
	bStateSafe:=FALSE;
END_IF
rtStateSafe(CLK:=bStateSafe);
ftStateSafe(CLK:=bStateSafe);

IF bStateSafe THEN
	sBitmap_ESButton:= 'ImagePool.EStop_OK2';
	stBitMap:='bitmap\EStop_OK2.bmp';
ELSE
	sBitmap_ESButton:= 'ImagePool.EStop_ACT2';
	stBitMap:='bitmap\EStop_ACT2.bmp';
END_IF

(*
ton_TSafe_OK(IN:=g_IO.TSafeIn.InRun AND NOT g_IO.TSafeIn.COM_Err, PT:=T#1S );
IF ton_TSafe_OK.Q THEN;
	bStateSafe:=TRUE;
ELSE;
	bStateSafe:=FALSE;	
END_IF
rt_TSafe_OK(CLK:=ton_TSafe_OK.Q );
IF rt_TSafe_OK.Q THEN;
	m_Print_Success_Message();
END_IF



rt_TSafe_Err(CLK:=g_IO.TSafeIn.COM_Err);
IF rt_TSafe_Err.Q THEN;
	m_Print_Error_Message();
END_IF

ton_TSafe_Err_Reset_ON(IN:=g_IO.TSafeIn.COM_Err AND NOT g_IO.TSafeOut.ErrACK, PT:=T#2S );
IF ton_TSafe_Err_Reset_ON.Q THEN;
	g_IO.TSafeOut.ErrACK:=TRUE;
END_IF

ton_TSafe_Err_Reset_OFF(IN:=g_IO.TSafeOut.ErrACK, PT:=T#1S );
IF ton_TSafe_Err_Reset_OFF.Q THEN;
	g_IO.TSafeOut.ErrACK:=FALSE;
END_IF
*)

ACTION act_Call_TSs:
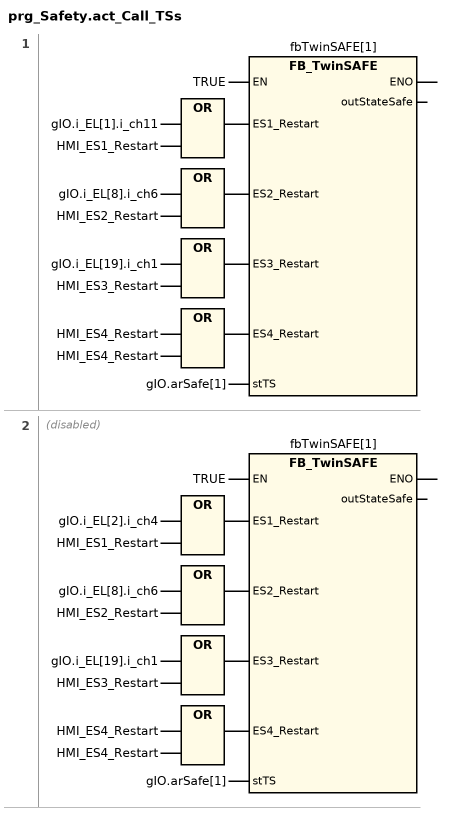
// NETWORK 1
fbTwinSAFE[1](
    ES1_Restart := gIO.i_EL[1].i_ch11 OR HMI_ES1_Restart,
    ES2_Restart := gIO.i_EL[8].i_ch6 OR HMI_ES2_Restart,
    ES3_Restart := gIO.i_EL[19].i_ch1 OR HMI_ES3_Restart,
    ES4_Restart := HMI_ES4_Restart OR HMI_ES4_Restart,
    stTS := gIO.arSafe[1]); // FB_TwinSAFE

// NETWORK 2 (disabled)
// fbTwinSAFE[1](
//     ES1_Restart := gIO.i_EL[2].i_ch4 OR HMI_ES1_Restart,
//     ES2_Restart := gIO.i_EL[8].i_ch6 OR HMI_ES2_Restart,
//     ES3_Restart := gIO.i_EL[19].i_ch1 OR HMI_ES3_Restart,
//     ES4_Restart := HMI_ES4_Restart OR HMI_ES4_Restart,
//     stTS := gIO.arSafe[1]); // FB_TwinSAFE
END_ACTION

METHOD m_Print_Error_Message : BOOL
VAR_INPUT
END_VAR

VAR
	i: INT;
	sActErrorID: STRING(11);
	sModuleDescription: STRING(80);
END_VAR

sActErrorID:='0x999x0';
sModuleDescription:='TwinSAFE Group';

FOR i:=100 TO 2 BY -1 DO
	Buffer_Act_Message[i]:=Buffer_Act_Message[i-1];
END_FOR

Buffer_Act_Message[1].sDateTime:=sRealTime_Date;
Buffer_Act_Message[1].sErrID:=sActErrorID;
Buffer_Act_Message[1].sModuleDescription:=sModuleDescription;
Buffer_Act_Message[1].sLevel:='Error';
Buffer_Act_Message[1].sErrorMessage:='';

Buffer_Act_Message[1].sErrorMessage:=CONCAT(Buffer_Act_Message[1].sErrorMessage,'TwinSAFE group has a communication error');
FUN_Write_Line_To_History();
END_METHOD

METHOD m_Print_Success_Message : BOOL
VAR_INPUT
END_VAR

VAR
	i: INT;
	sActErrorID: STRING(11);
	sModuleDescription: STRING(80);
END_VAR

sActErrorID:='0x999x0';
sModuleDescription:='TwinSAFE Group';

FOR i:=1000 TO 2 BY -1 DO
	Buffer_Act_History[i]:=Buffer_Act_History[i-1];
END_FOR

Buffer_Act_History[1].sDateTime:=sRealTime_Date;
Buffer_Act_History[1].sErrID:=sActErrorID;
Buffer_Act_History[1].sModuleDescription:=sModuleDescription;
Buffer_Act_History[1].sLevel:='Message';
Buffer_Act_History[1].sErrorMessage:='';

Buffer_Act_History[1].sErrorMessage:=CONCAT(Buffer_Act_History[1].sErrorMessage,'TwinSAFE state is OK');
END_METHOD

END_PROGRAM

// ---- 00 Library/05 Safety/FB_TwinSAFE.TcPOU
FUNCTION_BLOCK FB_TwinSAFE
VAR_INPUT
	ES1_Restart: BOOL;
	ES2_Restart: BOOL;
	ES3_Restart: BOOL;
	ES4_Restart: BOOL;
END_VAR
VAR_OUTPUT
	outStateSafe: BOOL;
END_VAR
VAR
	rt_TSafe_OK: R_TRIG;
	rt_TSafe_Err: R_TRIG;
	ton_TSafe_OK: TON;
	ton_TSafe_Err_Reset_ON: TON;
	ton_TSafe_Err_Reset_OFF: TON;	
END_VAR
VAR_IN_OUT
	stTS: ST_TwinSAFE;
END_VAR

stTS.stSafetyOut.ES1_PB_Restart:=ES1_Restart;
stTS.stSafetyOut.ES2_PB_Restart:=ES2_Restart;
stTS.stSafetyOut.ES3_PB_Restart:=ES3_Restart;
stTS.stSafetyOut.ES4_PB_Restart:=ES4_Restart;


//stTS.TSafeOut.Restart:=ES1_Restart;

ton_TSafe_OK(IN:=stTS.TSafeIn.InRun AND NOT stTS.TSafeIn.COM_Err, PT:=T#1S );
IF ton_TSafe_OK.Q 
AND stTS.stSafetyIn.ES1_State
AND stTS.stSafetyIn.ES2_State
AND stTS.stSafetyIn.ES3_State
AND stTS.stSafetyIn.ES4_State
THEN;
	outStateSafe:=TRUE;
ELSE;
	outStateSafe:=FALSE;	
END_IF
rt_TSafe_OK(CLK:=ton_TSafe_OK.Q );
IF rt_TSafe_OK.Q THEN;
	//m_Print_Success_Message();
END_IF



rt_TSafe_Err(CLK:=stTS.TSafeIn.COM_Err);
IF rt_TSafe_Err.Q THEN;
	//m_Print_Error_Message();
END_IF

ton_TSafe_Err_Reset_ON(IN:=stTS.TSafeIn.COM_Err AND NOT stTS.TSafeOut.ErrACK, PT:=T#2S );
IF ton_TSafe_Err_Reset_ON.Q THEN;
	stTS.TSafeOut.ErrACK:=TRUE;
END_IF

ton_TSafe_Err_Reset_OFF(IN:=stTS.TSafeOut.ErrACK, PT:=T#1S );
IF ton_TSafe_Err_Reset_OFF.Q THEN;
	stTS.TSafeOut.ErrACK:=FALSE;
END_IF

METHOD m_Print_Error_Message : BOOL
VAR_INPUT
END_VAR

VAR
	i: INT;
	sActErrorID: STRING(11);
	sModuleDescription: STRING(80);
END_VAR

sActErrorID:='0x999x0';
sModuleDescription:='TwinSAFE Group';

FOR i:=100 TO 2 BY -1 DO
	Buffer_Act_Message[i]:=Buffer_Act_Message[i-1];
END_FOR

Buffer_Act_Message[1].sDateTime:=sRealTime_Date;
Buffer_Act_Message[1].sErrID:=sActErrorID;
Buffer_Act_Message[1].sModuleDescription:=sModuleDescription;
Buffer_Act_Message[1].sLevel:='Error';
Buffer_Act_Message[1].sErrorMessage:='';

Buffer_Act_Message[1].sErrorMessage:=CONCAT(Buffer_Act_Message[1].sErrorMessage,'TwinSAFE group has a communication error');
FUN_Write_Line_To_History();
END_METHOD

METHOD m_Print_Success_Message : BOOL
VAR_INPUT
END_VAR

VAR
	i: INT;
	sActErrorID: STRING(11);
	sModuleDescription: STRING(80);
END_VAR

sActErrorID:='0x999x0';
sModuleDescription:='TwinSAFE Group';

FOR i:=1000 TO 2 BY -1 DO
	Buffer_Act_History[i]:=Buffer_Act_History[i-1];
END_FOR

Buffer_Act_History[1].sDateTime:=sRealTime_Date;
Buffer_Act_History[1].sErrID:=sActErrorID;
Buffer_Act_History[1].sModuleDescription:=sModuleDescription;
Buffer_Act_History[1].sLevel:='Message';
Buffer_Act_History[1].sErrorMessage:='';

Buffer_Act_History[1].sErrorMessage:=CONCAT(Buffer_Act_History[1].sErrorMessage,'TwinSAFE state is OK');
END_METHOD

END_FUNCTION_BLOCK

// ---- 01 Instance/04-Messages/prg_MessageManager.TcPOU
PROGRAM prg_MessageManager
VAR
	i_count         : INT;
	i_Reset         : INT;

	i_Buffer        : INT;
	i_Index         : INT;
	rtPressostat    : R_TRIG;
	PressostatFilter: TON;
	i               : INT;
	bAirPressureOk  : BOOL;
	ton_Error_201_Delay: TON;
	ton_Error_202_Delay: TON;
	ton_Error_251_Delay: TON;
	ton_Error_252_Delay: TON;
	ton_Error_253_Delay: TON;
	ton_Error_203_Delay: TON;
	ton_Error_204_Delay: TON;
	c_Unknown     : INT;
	iNumber       : INT;
	sNumber       : STRING(4);
	iNumber2      : INT;
	sNumber2      : STRING(4);
	iNumber4      : INT;
	sNumber4      : STRING(4);
	iNumber5      : INT;
	sNumber5      : STRING(4);
	rt_Print: R_TRIG;
	sModuleID: STRING(3);
	sModuleDescriptionHMI: STRING;
	testMessage: BOOL;
END_VAR

VAR_INPUT
	b_ResetAll    : BOOL;
END_VAR

prg_MessageManager.act_Count();
prg_MessageManager.act_GeneralMessage();
prg_MessageManager.act_Tanks_Lock();
//prg_MessageManager.act_AirPressure();

 m_AirPressure(aSense_Name:=E_ASense_Name.AP1001);
 //Zones 2..4 (TriBlender, Marinade, Color) are not used by the local CIP
 //m_AirPressure(aSense_Name:=E_ASense_Name.AP2001);
 //m_AirPressure(aSense_Name:=E_ASense_Name.AP3001);
 //m_AirPressure(aSense_Name:=E_ASense_Name.AP4001);

 // Motors
m_Motor(ePump_name:=E_Pump_List.P1001);
//m_Motor(ePump_name:=E_Pump_List.P3001);
//m_Motor(ePump_name:=E_Pump_List.P3002);
//m_Motor(ePump_name:=E_Pump_List.AG3001);
//m_Motor(ePump_name:=E_Pump_List.AG3002);
//m_Motor(ePump_name:=E_Pump_List.P4001);
//m_Motor(ePump_name:=E_Pump_List.P4002);
//m_Motor(ePump_name:=E_Pump_List.AG4001);
//m_Motor(ePump_name:=E_Pump_List.AG4002);
//m_Motor(ePump_name:=E_Pump_List.TB0001);

ACTION act_AirPressure:

 m_AirPressure(aSense_Name:=E_ASense_Name.AP1001);
 m_AirPressure(aSense_Name:=E_ASense_Name.AP2001);
 m_AirPressure(aSense_Name:=E_ASense_Name.AP3001);
 m_AirPressure(aSense_Name:=E_ASense_Name.AP4001);
END_ACTION

ACTION act_Count:
	iActErrors:=0;
	iActMessages:=0;
	iActWarning:=0;
FOR i_count:=1 TO 100 BY 1 DO

	IF Buffer_Act_Message[i_count].sLevel<>'' THEN
		IF Buffer_Act_Message[i_count].sLevel='Error' THEN
			iActErrors:=iActErrors+1;
		ELSIF Buffer_Act_Message[i_count].sLevel='Warning' OR Buffer_Act_Message[i_count].sLevel='Error temp'THEN
			iActWarning:=iActWarning+1;
		ELSIF Buffer_Act_Message[i_count].sLevel='Message' THEN
			iActMessages:=iActMessages+1;		
		END_IF
	END_IF

END_FOR
END_ACTION

ACTION act_GeneralMessage:
;
			(*-------------------->Air Pressure<--------------------*)
	bAirPressureOk:= TRUE;  //i_EP[18].x0
	IF   NOT bAirPressureOk THEN //bAirPressureSensorExist AND
		//ar_Message[1].b_Active:=TRUE;	(*	Air_Pressure_Too_Low	*)
		fbPrintErrMessageByID(sModuleDescription:='General',sActErrorID:='050x000x001');
	ELSE;
		//ar_Message[1].b_Active:=FALSE;	(*	Air_Pressure_Too_Low	*)
	END_IF








			(*-------------------->Emergency<--------------------*)
	IF bES_Bypass THEN;
		//'106x000x060',   'Warning',    'Emergency Bypass activated,	
		fbPrintErrMessageByID(sModuleDescription:='Emergency',sActErrorID:='106x000x060');
	ELSE;	
		//IF NOT bStateSafe THEN
		
		IF NOT arSafe[1].stSafetyIn.ES1_State THEN
			fbPrintErrMessageByID(sModuleDescription:='Emergency 1',sActErrorID:='106x001x001');
		END_IF
		
// 		IF NOT arSafe[1].stSafetyIn.ES2_State THEN
// 			fbPrintErrMessageByID(sModuleDescription:='Emergency 2',sActErrorID:='106x002x001');
// 		END_IF		
		
		IF NOT arSafe[1].stSafetyIn.ES3_State THEN
			fbPrintErrMessageByID(sModuleDescription:='Emergency 3',sActErrorID:='106x003x001');			
		END_IF	
	
// 		IF NOT arSafe[1].stSafetyIn.ES4_State THEN
// 			fbPrintErrMessageByID(sModuleDescription:='Emergency 4',sActErrorID:='106x004x001');
// 		END_IF
		
		
		//IF NOT bES_PB[1].State THEN
		IF NOT arSafe[1].stSafetyIn.ES1_PB_State THEN
			fbPrintErrMessageByID(sModuleDescription:='Emergency 1',sActErrorID:='106x001x002');
		END_IF
// 		IF NOT arSafe[1].stSafetyIn.ES2_PB_State THEN
// 			fbPrintErrMessageByID(sModuleDescription:='Emergency 2',sActErrorID:='106x002x002');
// 		END_IF
		IF NOT arSafe[1].stSafetyIn.ES3_PB1_State THEN
			fbPrintErrMessageByID(sModuleDescription:='Emergency 3',sActErrorID:='106x003x002');
		END_IF
		IF NOT arSafe[1].stSafetyIn.ES3_PB2_State THEN
			fbPrintErrMessageByID(sModuleDescription:='Emergency 3',sActErrorID:='106x003x003');
		END_IF		
// 		IF NOT arSafe[1].stSafetyIn.ES4_PB_State THEN
// 			fbPrintErrMessageByID(sModuleDescription:='Emergency 4',sActErrorID:='106x004x002');
// 		END_IF
		
	END_IF
	
//test
		IF testMessage THEN
			fbPrintErrMessageByID(sModuleDescription:='eTank1',sActErrorID:='000x000x999');
		END_IF	
			(*-------------------->Doors Closed<--------------------*)
	(*
	IF NOT bInterlock[1] THEN;
		ar_Message[1].b_Active:=TRUE;
		fbPrintErrMessageByID(sModuleDescription:='Doors',sActErrorID:='107x000x101');
	ELSE
		IF NOT bInterlock[2] THEN;
			ar_Message[2].b_Active:=TRUE;
			fbPrintErrMessageByID(sModuleDescription:='Doors',sActErrorID:='107x000x102');
		ELSE
			IF NOT bInterlock[3] THEN;
				ar_Message[3].b_Active:=TRUE;
				fbPrintErrMessageByID(sModuleDescription:='Doors',sActErrorID:='107x000x103');
			ELSE				
				ar_Message[3].b_Active:=FALSE;
			END_IF					
			ar_Message[2].b_Active:=FALSE;
		END_IF			
		ar_Message[1].b_Active:=FALSE;
	END_IF	
	*)
	(*		
	FOR i:=4 TO 8 DO
		IF NOT bInterlock[i] THEN
			ar_Message[100+i].b_Active:=TRUE;	(*	Door_Num_1_Not_Closed	*)
			iNumber := 100+i;
			sNumber := INT_TO_STRING (iNumber);
			
		ELSE
			ar_Message[100+i].b_Active:=FALSE;
		END_IF
	END_FOR
	*)
			(*-------------------->Doors Locked<--------------------*)
			
	FOR i:=1 TO 12 DO
		iNumber2 := 120+i;
		sNumber2 := INT_TO_STRING (iNumber2);		
		CASE i OF 
			//Zone1 
			1,2,6,7:;
				IF bReq_LockZone[1] AND NOT bDoorLocked[i] THEN
					fbPrintErrMessageByID(sModuleDescription:='Doors',sActErrorID:=concat ('107x000x', sNumber2));
				END_IF	
		END_CASE
		CASE i OF 		
			//Zone2
			2,3,4:;
				IF bReq_LockZone[2] AND NOT bDoorLocked[i] THEN
					fbPrintErrMessageByID(sModuleDescription:='Doors',sActErrorID:=concat ('107x000x', sNumber2));
				END_IF	
		END_CASE
		CASE i OF 			
			//Zone3
			5,6:;
				IF bReq_LockZone[3] AND NOT bDoorLocked[i] THEN
					fbPrintErrMessageByID(sModuleDescription:='Doors',sActErrorID:=concat ('107x000x', sNumber2));
				END_IF		
		END_CASE
		CASE i OF 					
			//Zone4
			3,4,5:;
				IF bReq_LockZone[4] AND NOT bDoorLocked[i] THEN
					fbPrintErrMessageByID(sModuleDescription:='Doors',sActErrorID:=concat ('107x000x', sNumber2));
				END_IF							
			
		END_CASE

	END_FOR
	
	
			(*-------------------->Intrlock Zones<--------------------*)
	FOR i:=1 TO 4 DO
		IF bReq_LockZone[1] AND (NOT bIntZoneLocked[i]) AND (NOT bIntZoneBypass[i]) THEN
			iNumber4 := 140+i;
			sNumber4 := INT_TO_STRING (iNumber4);
			fbPrintErrMessageByID(sModuleDescription:='Inter lock Zone',sActErrorID:=concat ('108x000x', sNumber4));
		END_IF
	END_FOR
END_ACTION

ACTION act_Tanks_Lock:
{IF defined (Production)}
	IF NOT gIO.arSafe[1].stSafetyIn.TankLocked_CIP_T91 THEN
		fbPrintErrMessageByID(sModuleDescription:='Tank Interlock',sActErrorID:='101x002xT91');
	END_IF
	IF NOT gIO.arSafe[1].stSafetyIn.TankLocked_CIP_T92 THEN
		fbPrintErrMessageByID(sModuleDescription:='Tank Interlock',sActErrorID:='101x002xT92');
	END_IF
	IF NOT gIO.arSafe[1].stSafetyIn.TankLocked_CIP_T93 THEN
		fbPrintErrMessageByID(sModuleDescription:='Tank Interlock',sActErrorID:='101x002xT93');
	END_IF
	IF NOT gIO.arSafe[1].stSafetyIn.TankLocked_CIP_T94 THEN
		fbPrintErrMessageByID(sModuleDescription:='Tank Interlock',sActErrorID:='101x002xT94');
	END_IF
	
// 	IF NOT gIO.arSafe[1].stSafetyIn.TankLocked_Marinade_T1 THEN
// 		//fbPrintErrMessageByID(sModuleDescription:='Tank Interlock',sActErrorID:='101x002xT01');
// 	END_IF
// 	IF NOT gIO.arSafe[1].stSafetyIn.TankLocked_Marinade_T2 THEN
// 		//fbPrintErrMessageByID(sModuleDescription:='Tank Interlock',sActErrorID:='101x002xT02');
// 	END_IF
	
// 	IF NOT gIO.arSafe[1].stSafetyIn.TankLocked_Color_T3 THEN
// 		fbPrintErrMessageByID(sModuleDescription:='Tank Interlock',sActErrorID:='101x002xT03');
// 	END_IF
// 	IF NOT gIO.arSafe[1].stSafetyIn.TankLocked_Color_T4 THEN
// 		fbPrintErrMessageByID(sModuleDescription:='Tank Interlock',sActErrorID:='101x002xT04');
// 	END_IF
{ELSIF defined (Simulation_IO)}
{END_IF}
END_ACTION

METHOD m_AirPressure : BOOL
VAR_INPUT
	aSense_Name: E_ASense_Name;
END_VAR

VAR
	k: STRING(1);
	temp_string: STRING(3);
END_VAR

{IF defined (Production)}
	IF TRUE
	//AND __ISVALIDREF(fbAnalogSensor[aSense_Name]) 
	THEN;
		
		temp_string:=TO_STRING(aSense_Name);
		k:=MID(temp_string, 3, 3);
		
		IF fbAnalogSensor[aSense_Name].bLL_Warning THEN;
			fbPrintErrMessageByID(sModuleDescription:='Air Pressure',sActErrorID:=concat ('101x003x01', k));
		END_IF
		
		IF fbAnalogSensor[aSense_Name].bHH_Warning THEN;
			fbPrintErrMessageByID(sModuleDescription:='Air Pressure',sActErrorID:=concat ('101x003x02', k));
		END_IF
		
		IF fbAnalogSensor[aSense_Name].bLL_Alarm THEN;
			fbPrintErrMessageByID(sModuleDescription:='Air Pressure',sActErrorID:=concat ('101x003x11', k));
		END_IF
		
		IF fbAnalogSensor[aSense_Name].bHH_Alarm THEN;
			fbPrintErrMessageByID(sModuleDescription:='Air Pressure',sActErrorID:=concat ('101x003x12', k));
		END_IF
		
		
	ELSE;
		RETURN;
	END_IF
{ELSIF defined (Simulation_IO)}
{END_IF}
END_METHOD

METHOD m_Motor : BOOL
VAR_INPUT
	ePump_name: E_Pump_List;
END_VAR

VAR
	temp_string: STRING(6);
END_VAR
{IF defined (Production)}
temp_string:=TO_STRING(ePump_name);

IF g_Pump.fbPump[ePump_name].m_Error()<>'' THEN;
	fbPrintErrMessageByID(sModuleDescription:='Motor', sActErrorID:=g_Pump.fbPump[ePump_name].m_Error());
END_IF
{ELSIF defined (Simulation_IO)}
{END_IF}
END_METHOD

END_PROGRAM

// ---- 01 Instance/04-Messages/prg_Messages.TcPOU
PROGRAM prg_Messages
VAR
	Pis: INT;
	c_PisError: INT;
	mask_PisEr: ARRAY [1..C_Max_Pistons] OF BOOL;
	mask_LatEr: ARRAY [1..24] OF BOOL;
	Mess: INT;
	ResetErrors: BOOL;
	(*ResumeAll: BOOL;*)
	r_trig_prg_Stepper: R_TRIG;
	r_trig_StepperErrorSFC: R_TRIG;
	ton_ActMessCheck: TON;
	sel_FB: INT;
	PauseAll: BOOL;
	Lat: INT;

	HighLightErrorPB: BOOL;
	HighLightWarningPB: BOOL;
	
	Clear: STRING := '';
	ton_BitMapBlink: TON;
	stBitMap: STRING;
	r_trig_ResetError: R_trig;
	i_Reset: INT;
END_VAR

ton_ActMessCheck(IN:=NOT ton_ActMessCheck.Q, PT:=T#0.5S);

prg_Messages.act_ResetErrors();
prg_Messages.act_ResumeSFC();


IF iActErrors<>0 THEN
	HighLightErrorPB:=TRUE;
ELSE
	HighLightErrorPB:=FALSE;
END_IF

IF iActWarning<>0 THEN
	HighLightWarningPB:=TRUE;
ELSE
	HighLightWarningPB:=FALSE;
END_IF

ton_BitMapBlink(PT:=T#1S,IN:=NOT ton_BitMapBlink.Q);
IF HighLightErrorPB THEN
	IF ton_BitMapBlink.ET>T#0.5S THEN
		 s_Error_BitmapID:='ImagePool.Error_Yel';
	ELSE
		 s_Error_BitmapID:='ImagePool.Error_Red';
	END_IF
ELSIF HighLightWarningPB THEN
	IF ton_BitMapBlink.ET>T#0.5S THEN
		 s_Error_BitmapID:='ImagePool.Error_Yel';
	ELSE
		 s_Error_BitmapID:='ImagePool.Error_No';
	END_IF
ELSE
		 s_Error_BitmapID:='ImagePool.Error_No';
END_IF

ACTION act_ResetErrors:
r_trig_ResetError(CLK:=ResetErrors OR
						stOpMain.bResetError );

IF r_trig_ResetError.Q THEN
	(*	 Pistons		*)
	FOR Pis:=1 TO C_Max_Pistons BY 1 DO
		stPis[Pis].b_Resume:=TRUE;
	END_FOR
	FOR i_Reset:=1 TO 100 BY 1 DO
		Buffer_Act_Message[i_Reset].sDateTime:='';
		Buffer_Act_Message[i_Reset].sErrID:='';
		Buffer_Act_Message[i_Reset].sLevel:='';
		Buffer_Act_Message[i_Reset].sErrorMessage:='';
		Buffer_Act_Message[i_Reset].sModuleDescription:='';
	END_FOR
END_IF

IF ResetErrors THEN

(*		 Pistons		*)
	FOR Pis:=1 TO C_Max_Pistons BY 1 DO
		stPis[Pis].b_Resume:=TRUE;
	END_FOR

(*		Latches		*)
	(*FOR Pis:=1 TO 24 BY 1 DO
		db_Lat[Pis].req_Resume:=TRUE;
	END_FOR*)

	//prg_Safety.ResetError:=TRUE;

	ResetErrors:=FALSE;
END_IF
END_ACTION

ACTION act_ResumeSFC:
IF ResumeAll THEN

(*		 Pistons		*)
	FOR Pis:=1 TO C_Max_Pistons BY 1 DO
		stPis[Pis].b_Resume:=TRUE;
	END_FOR


(*		Latches		*)
	(*FOR Pis:=1 TO 24 BY 1 DO
		db_Lat[Pis].req_Resume:=TRUE;
	END_FOR*)



	ResetErrors:=TRUE;
END_IF
END_ACTION

END_PROGRAM

// ---- 01 Instance/07-Mode/prg_Call_OpMode.TcPOU
PROGRAM prg_Call_OpMode
VAR
	fbModeMain:FB_ModeSelect;
	
	rt_HMI_Resume: R_TRIG;
	rt_ActError: R_TRIG;
	
	eModeZone: E_ModeZone;

END_VAR

fbModeMain(sModuleDescription:='Mode Select - Main',
	bInterlockBypass:=TRUE, //bIntZoneBypass[1]
	bLockedFB:=TRUE, //bIntZoneLocked[1]
	bPistonCheck:=FALSE,	
	bLockRequest=>,	//bReq_LockZone[1]
	eModeZone:=E_ModeZone.eMain,
	stMode:=stModeMain,
	stOperation:=stOpMain, 
	bStateSafe_mode:=bStateSafe);
	
FOR eModeZone:=	E_ModeZone.eMain TO E_ModeZone.eLast DO
	fbMode[eModeZone](sModuleDescription:='Mode Select - ',
		bInterlockBypass:=TRUE, //bIntZoneBypass[eModeZone]
		bLockedFB:=TRUE, //bIntZoneLocked[eModeZone]
		bPistonCheck:=FALSE,	
		bLockRequest=>,	//bReq_LockZone[eModeZone]
		eModeZone:=eModeZone,
		stMode:=stMode[eModeZone],
		stOperation:=stOper[eModeZone],
		bStateSafe_mode:=m_Get_StateSafe_by_ModeZone(eMoZone:=eModeZone));	
END_FOR
	
PauseAll:=stOpMain.iActOperation=E_OperationButtons.ePauseAll;	
PauseAllDelayed:=stOpMain.bPauseOnDelayed;	

stOpNonPause.iActOperation:=E_OperationButtons.ePlayAll;
	
rt_HMI_Resume(CLK:=ResumeAll);
IF rt_HMI_Resume.Q THEN;
	stOpMain.bSetPlay:=TRUE;
	prg_Messages.act_ResumeSFC();	
	FOR eModeZone:=	E_ModeZone.eMain TO E_ModeZone.eLast DO;
		stOper[eModeZone].bSetPlay:=TRUE;
	END_FOR
END_IF
ResumeAll:=FALSE;

rt_ActError(CLK:=iActErrors<>0);
IF iActErrors<>0 THEN;
	stOpMain.bSetPause:=TRUE;
END_IF

prg_LightTower(
	bBuzzerBypass:=bBuzzerMute , 
	qLedGreen=> , //q_EL16[2].ch11
	qLedYellow=> , //q_EL16[2].ch10
	qLedRed=> , //q_EL16[2].ch9
	qBuzzer=> );//q_EL16[2].ch12
	
	
act_Call_LightTowers();

ACTION act_Call_LightTowers:
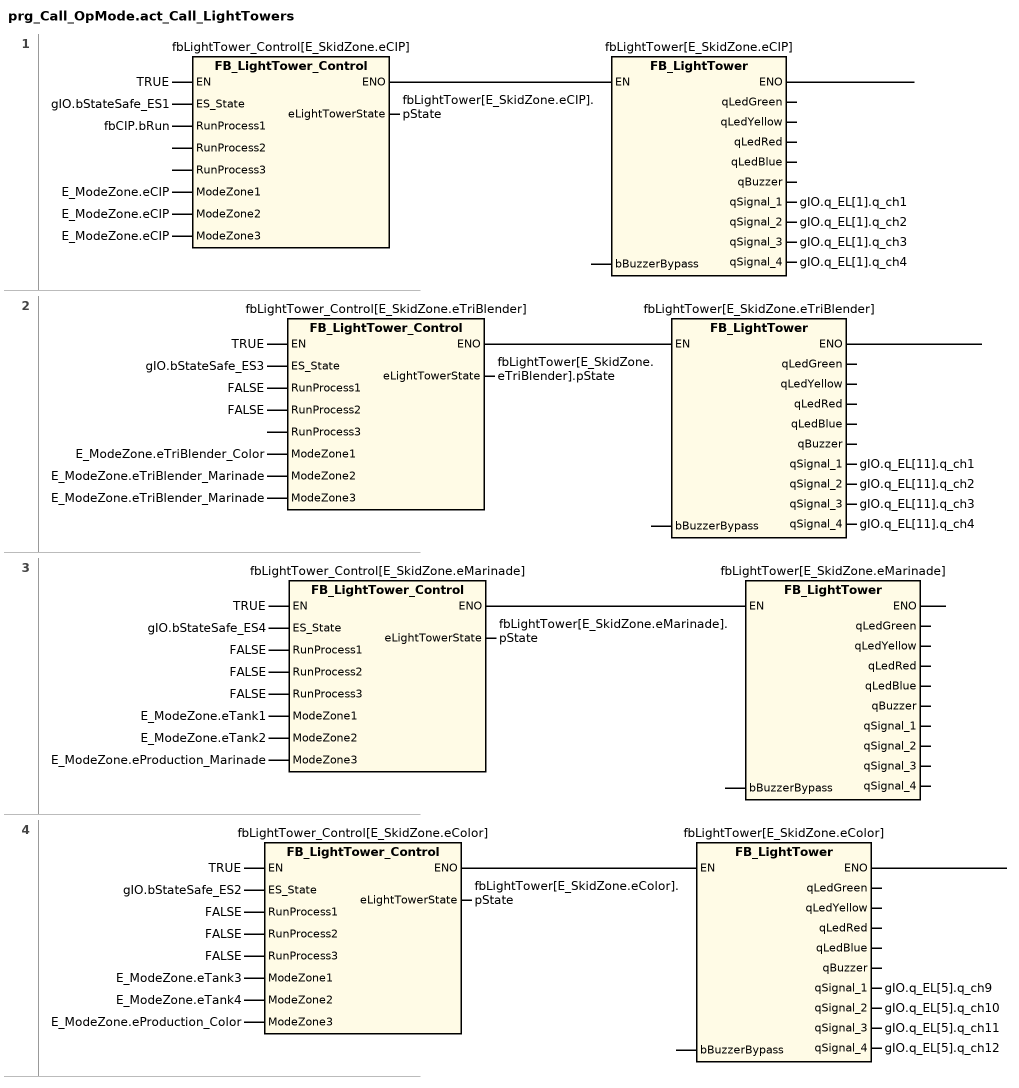
// NETWORK 1
fbLightTower_Control[E_SkidZone.eCIP](
    ES_State := gIO.bStateSafe_ES1,
    RunProcess1 := fbCIP.bRun,
    ModeZone1 := E_ModeZone.eCIP,
    ModeZone2 := E_ModeZone.eCIP,
    ModeZone3 := E_ModeZone.eCIP,
    eLightTowerState => fbLightTower[E_SkidZone.eCIP].pState); // FB_LightTower_Control
fbLightTower[E_SkidZone.eCIP](
    qSignal_1 => gIO.q_EL[1].q_ch1,
    qSignal_2 => gIO.q_EL[1].q_ch2,
    qSignal_3 => gIO.q_EL[1].q_ch3,
    qSignal_4 => gIO.q_EL[1].q_ch4); // FB_LightTower

// NETWORK 2
fbLightTower_Control[E_SkidZone.eTriBlender](
    ES_State := gIO.bStateSafe_ES3,
    RunProcess1 := FALSE,
    RunProcess2 := FALSE,
    ModeZone1 := E_ModeZone.eTriBlender_Color,
    ModeZone2 := E_ModeZone.eTriBlender_Marinade,
    ModeZone3 := E_ModeZone.eTriBlender_Marinade,
    eLightTowerState => fbLightTower[E_SkidZone.eTriBlender].pState); // FB_LightTower_Control
fbLightTower[E_SkidZone.eTriBlender](
    qSignal_1 => gIO.q_EL[11].q_ch1,
    qSignal_2 => gIO.q_EL[11].q_ch2,
    qSignal_3 => gIO.q_EL[11].q_ch3,
    qSignal_4 => gIO.q_EL[11].q_ch4); // FB_LightTower

// NETWORK 3
fbLightTower_Control[E_SkidZone.eMarinade](
    ES_State := gIO.bStateSafe_ES4,
    RunProcess1 := FALSE,
    RunProcess2 := FALSE,
    RunProcess3 := FALSE,
    ModeZone1 := E_ModeZone.eTank1,
    ModeZone2 := E_ModeZone.eTank2,
    ModeZone3 := E_ModeZone.eProduction_Marinade,
    eLightTowerState => fbLightTower[E_SkidZone.eMarinade].pState); // FB_LightTower_Control
fbLightTower[E_SkidZone.eMarinade](); // FB_LightTower

// NETWORK 4
fbLightTower_Control[E_SkidZone.eColor](
    ES_State := gIO.bStateSafe_ES2,
    RunProcess1 := FALSE,
    RunProcess2 := FALSE,
    RunProcess3 := FALSE,
    ModeZone1 := E_ModeZone.eTank3,
    ModeZone2 := E_ModeZone.eTank4,
    ModeZone3 := E_ModeZone.eProduction_Color,
    eLightTowerState => fbLightTower[E_SkidZone.eColor].pState); // FB_LightTower_Control
fbLightTower[E_SkidZone.eColor](
    qSignal_1 => gIO.q_EL[5].q_ch9,
    qSignal_2 => gIO.q_EL[5].q_ch10,
    qSignal_3 => gIO.q_EL[5].q_ch11,
    qSignal_4 => gIO.q_EL[5].q_ch12); // FB_LightTower
END_ACTION

METHOD INTERNAL m_Get_StateSafe_by_ModeZone : BOOL
VAR_INPUT
	eMoZone: E_ModeZone;
END_VAR
CASE eMoZone OF
	E_ModeZone.eCIP:;
		m_Get_StateSafe_by_ModeZone:=bStateSafe_ES1;

	E_ModeZone.eTank3,
	E_ModeZone.eTank4,
	E_ModeZone.eProduction_Color:;
		m_Get_StateSafe_by_ModeZone:=bStateSafe_ES2;		

	E_ModeZone.eTriBlender_Color,
	E_ModeZone.eTriBlender_Marinade:;
		m_Get_StateSafe_by_ModeZone:=bStateSafe_ES3;
		
	E_ModeZone.eTank1,
	E_ModeZone.eTank2,
	E_ModeZone.eProduction_Marinade:;
		m_Get_StateSafe_by_ModeZone:=bStateSafe_ES4;
		
ELSE;
		m_Get_StateSafe_by_ModeZone:=FALSE;
		
END_CASE
(*
bStateSafe_ES1:=arSafe[1].stSafetyIn.ES1_State;
bStateSafe_ES2:=arSafe[1].stSafetyIn.ES2_State;
bStateSafe_ES3:=arSafe[1].stSafetyIn.ES3_State;
bStateSafe_ES4:=arSafe[1].stSafetyIn.ES4_State;
*)
END_METHOD

END_PROGRAM

// ---- 00 Library/07-Mode/FB_ModeSelect.TcPOU
FUNCTION_BLOCK FB_ModeSelect
VAR_INPUT
	bInterlockBypass: BOOL;
	bAutoPlayEnable: BOOL:=TRUE;
	sModuleDescription: STRING:='Mode Select';
	eModeZone:E_ModeZone;
	bLockedFB: BOOL;
	bPistonCheck: BOOL:=TRUE;
	bStateSafe_mode: BOOL:=TRUE;
END_VAR
VAR_OUTPUT
	bModeStillState: BOOL;
	bLockRequest: BOOL;
END_VAR
VAR
	fbPrintErrMessageByID: FB_PrintErrMessageByID_SFC_Cycle;
	r_trig_ModeExchange1: R_TRIG;
	r_trig_ModeExchange2: R_TRIG;
	r_trig_ModeExchange3: R_TRIG;
	ton_ModeExchengeDelay: TON;	
	fbOperation:FB_Operation;
	bLockRelay: BOOL;	
	i: INT;
	bPistonsOK: BOOL;
	fbFormatString:FB_FormatString;
	sFB_ID: STRING(3):='050';

	sActErrorID: STRING(11);
	sFullErrorId: STRING(11);
	//r_trigAuto: R_TRIG;
	r_trigIntClose: R_TRIG;
	r_trigIntOpen: R_TRIG;
	bIntZonePaused: BOOL;
	rt_Play: R_TRIG;

END_VAR
VAR
	ton_ResumeMachine: TON;
	ton_ResetErrors: TON;
	ton_ResetAllCycles: TON;
	ton_PlayAllDelay: TON;
	ton_PauseDelay: TON;
	r_trigPlayAllDelay: R_TRIG;
	ton_PlayDelay: TON;
END_VAR
VAR_IN_OUT
	stMode:ST_Mode;
	stOperation:ST_OperationButtons;
END_VAR

act_Oper();
act_ModeStillState();
fbOperation(stOper:=stOperation);
stMode.eModeZone:=eModeZone;		
stOperation.eModeZone:=eModeZone;
stOperation.sModeZone:=TO_STRING(eModeZone);
IF (stMode.iActMode=E_WorkingMode.eAutoMode OR stMode.iActMode=E_WorkingMode.eSemiAutoMode)
AND NOT bInterlockBypass
THEN;
	bLockRequest:=TRUE;
ELSE;
	bLockRequest:=FALSE;
END_IF



r_trigIntClose(CLK:=bLockedFB);
r_trigIntOpen(CLK:=NOT bLockedFB);

(*888888888888888888   InterLocks Zone 1		8888888888888*)
IF stOperation.iActOperation=E_OperationButtons.ePlayAll AND  r_trigIntOpen.Q THEN
	bIntZonePaused:=TRUE;
END_IF

IF NOT bLockedFB 
AND NOT bInterlockBypass	
AND stOperation.iActOperation=E_OperationButtons.ePlayAll THEN
	//Message
	sActErrorID:='351'; // '050x000x351',	'Warning',	'Interlock Paused Operation',
	act_GetErrorID_Format();
	fbPrintErrMessageByID(sFB_ModuleDescription:=sModuleDescription,sActErrorID:=sFullErrorId,bSFCError:=TRUE);
	stOperation.bSetPause:=TRUE;
	stOperation.iPauseHistory:=4;
END_IF


IF bAutoPlayEnable AND bIntZonePaused AND r_trigIntClose.Q THEN
	stOperation.bSetPlay:=TRUE;
	bIntZonePaused:=FALSE;
END_IF

IF bLockedFB OR stMode.iActMode=E_WorkingMode.eManualMode THEN
	bIntZonePaused:=FALSE;
END_IF

rt_Play(CLK:=stOperation.iActOperation=E_OperationButtons.ePlayAll);

IF NOT bStateSafe_mode OR stOperation.bStopResetAll THEN;
	stMode.bSetManual:=TRUE;
	stOperation.bSetPause:=TRUE;
END_IF

stMode.bStateSafe_mode:=stOperation.bStateSafe_mode:=bStateSafe_mode;

m_Error_zone_check();

stOperation.iActModeState:=stMode.iActMode;

ACTION act_AutomationLock_Failed:
sActErrorID:='306';//'050x000x306',	'Warning',	'Semi/Auto mode request rejected, automation lock failed',
act_GetErrorID_Format();
fbPrintErrMessageByID(sFB_ModuleDescription:=sModuleDescription,sActErrorID:=sFullErrorId,bSFCError:=TRUE);
END_ACTION

ACTION act_Done:
stMode.bSetManual:=FALSE;
stMode.bSetSemi:=FALSE;
stMode.bSetAuto:=FALSE;
//stMode.iErrorNum:=0;
//stMode.sErrorMessage:='No Error';
END_ACTION

ACTION act_GetErrorID_Format:
(*IF bErrorSFC THEN;
	
	IF    sLast_SFCErrorStep='WaitSenOpen' 							THEN sActErrorID:='001';
	ELSIF sLast_SFCErrorStep='WaitSenNotClose' 		   				THEN sActErrorID:='002';
	ELSIF sLast_SFCErrorStep='WaitSenClose' 						THEN sActErrorID:='003';
	ELSIF sLast_SFCErrorStep='WaitSenNotOpen' 						THEN sActErrorID:='004';
	ELSIF sLast_SFCErrorStep='No Status' 							THEN sActErrorID:='005';		
	ELSIF sLast_SFCErrorStep='No Valve Operation' 					THEN sActErrorID:='006';
	ELSIF sLast_SFCErrorStep='Not synchronized with cycle command' 	THEN sActErrorID:='007';
	ELSIF sLast_SFCErrorStep='SensorsChecking' 						THEN sActErrorID:='008';
	
	ELSE;
		 sActErrorID:='999';
	END_IF

ELSE
		 sActErrorID:='000';
END_IF*)

fbFormatString(
	sFormat:= '%.3sx%.3dx%.3s', 
	arg1:= F_STRINGEx(sFB_ID), 
	arg2:= F_INT(eModeZone), 
	arg3:= F_STRINGEx(sActErrorID), 
	sOut=>sFullErrorId );
END_ACTION

ACTION act_ModeStillState:

r_trig_ModeExchange1(CLK:=stMode.iActMode=eManualMode);
r_trig_ModeExchange2(CLK:=stMode.iActMode=eSemiAutoMode);
r_trig_ModeExchange3(CLK:=stMode.iActMode=eAutoMode);
ton_ModeExchengeDelay(PT:=T#0.5S);
(*IF ton_ModeExchengeDelay.Q THEN
	ton_ModeExchengeDelay.IN:=FALSE;
END_IF*)
IF r_trig_ModeExchange1.Q
OR r_trig_ModeExchange2.Q
OR r_trig_ModeExchange3.Q
THEN
	ton_ModeExchengeDelay(IN:=FALSE);
	ton_ModeExchengeDelay.IN:=TRUE;
END_IF
bModeStillState:=ton_ModeExchengeDelay.Q;
END_ACTION

ACTION act_Oper:
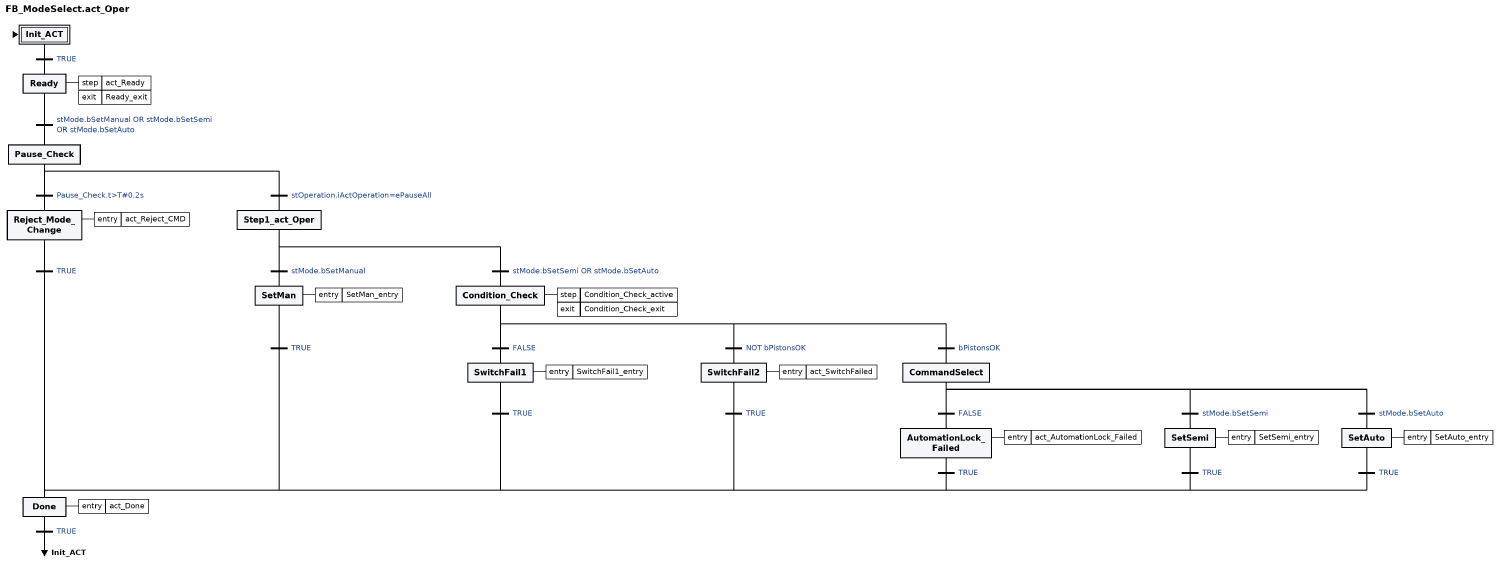
INITIAL_STEP Init_ACT:
END_STEP
TRANSITION FROM Init_ACT TO Ready
    := TRUE;
END_TRANSITION
STEP Ready:
    act_Ready(N);  // step action
    Ready_exit(P0);  // exit action
END_STEP
TRANSITION FROM Ready TO Pause_Check
    := stMode.bSetManual OR stMode.bSetSemi OR stMode.bSetAuto;
END_TRANSITION
STEP Pause_Check:
END_STEP
TRANSITION FROM Pause_Check TO Reject_Mode_Change
    := Pause_Check.t>T#0.2s;
END_TRANSITION
STEP Reject_Mode_Change:
    act_Reject_CMD(P1);  // entry action
END_STEP
TRANSITION FROM Reject_Mode_Change TO Done
    := TRUE;
END_TRANSITION
TRANSITION FROM Pause_Check TO Step1_act_Oper
    := stOperation.iActOperation=ePauseAll;
END_TRANSITION
STEP Step1_act_Oper:
END_STEP
TRANSITION FROM Step1_act_Oper TO SetMan
    := stMode.bSetManual;
END_TRANSITION
STEP SetMan:
    SetMan_entry(P1);  // entry action
END_STEP
TRANSITION FROM SetMan TO Done
    := TRUE;
END_TRANSITION
TRANSITION FROM Step1_act_Oper TO Condition_Check
    := stMode.bSetSemi OR stMode.bSetAuto;
END_TRANSITION
STEP Condition_Check:  // max time T#1s
    Condition_Check_active(N);  // step action
    Condition_Check_exit(P0);  // exit action
END_STEP
TRANSITION FROM Condition_Check TO SwitchFail1
    := FALSE;
END_TRANSITION
STEP SwitchFail1:
    SwitchFail1_entry(P1);  // entry action
END_STEP
TRANSITION FROM SwitchFail1 TO Done
    := TRUE;
END_TRANSITION
TRANSITION FROM Condition_Check TO SwitchFail2
    := NOT bPistonsOK;
END_TRANSITION
STEP SwitchFail2:
    act_SwitchFailed(P1);  // entry action
END_STEP
TRANSITION FROM SwitchFail2 TO Done
    := TRUE;
END_TRANSITION
TRANSITION FROM Condition_Check TO CommandSelect
    := bPistonsOK;
END_TRANSITION
STEP CommandSelect:  // max time T#1s
END_STEP
TRANSITION FROM CommandSelect TO AutomationLock_Failed
    := FALSE;
END_TRANSITION
STEP AutomationLock_Failed:
    act_AutomationLock_Failed(P1);  // entry action
END_STEP
TRANSITION FROM AutomationLock_Failed TO Done
    := TRUE;
END_TRANSITION
TRANSITION FROM CommandSelect TO SetSemi
    := stMode.bSetSemi;
END_TRANSITION
STEP SetSemi:
    SetSemi_entry(P1);  // entry action
END_STEP
TRANSITION FROM SetSemi TO Done
    := TRUE;
END_TRANSITION
TRANSITION FROM CommandSelect TO SetAuto
    := stMode.bSetAuto;
END_TRANSITION
STEP SetAuto:
    SetAuto_entry(P1);  // entry action
END_STEP
TRANSITION FROM SetAuto TO Done
    := TRUE;
END_TRANSITION
STEP Done:
    act_Done(P1);  // entry action
END_STEP
TRANSITION FROM Done TO Init_ACT
    := TRUE;
END_TRANSITION
// branch label Branch3_act_Oper
// branch label Branch1_act_Oper
// branch label Branch0_ACT
// branch label Branch2_act_Oper
END_ACTION

ACTION act_Operation:
(*
IF stOperation.bSetPlay THEN;
	bResumeMachine:=TRUE;
END_IF
ton_ResumeMachine(PT:=T#10MS,IN:=bResumeMachine,);
ton_PlayAllDelay(PT:=T#20MS);
IF ton_ResumeMachine.Q THEN;
	bResumeMachine:=FALSE;	
	stOperation.bSetPlay:=FALSE;
	ton_PlayAllDelay.IN:=TRUE;	
END_IF





r_trigPlayAllDelay(CLK:=ton_PlayAllDelay.Q);
IF r_trigPlayAllDelay.Q THEN	
	IF FALSE(*iActErrorNum=0*) THEN
		//stOperation.iActOperation:=E_OperationButtons.ePlayAll;
		stOperation.bSetPlay:=TRUE;
	END_IF	
END_IF


IF stOperation.bSetPause THEN;
	stOperation.iActOperation:=E_OperationButtons.ePauseAll;
	stOperation.bSetPause:=FALSE;
	ton_PlayAllDelay.IN:=FALSE;
END_IF



IF stOperation.iActOperation=E_OperationButtons.ePauseAll THEN;
	
ELSIF stOperation.iActOperation=E_OperationButtons.ePlayAll THEN;
	
END_IF

bPauseMachine:=stOperation.iActOperation=E_OperationButtons.ePauseAll;


ton_PauseDelay(PT:=T#1S, IN:=stOperation.iActOperation=E_OperationButtons.ePauseAll);
ton_PlayDelay(PT:=T#1S, IN:=stOperation.iActOperation=E_OperationButtons.ePlayAll);
*)
END_ACTION

ACTION act_Ready:

IF stMode.iActMode=eManualMode AND stMode.bSetManual THEN; stMode.bSetManual:=FALSE; END_IF
IF stMode.iActMode=eSemiAutoMode AND stMode.bSetSemi THEN; stMode.bSetSemi:=FALSE; END_IF

IF stMode.iActMode=eAutoMode 
AND stMode.bSetAuto THEN; 
	stMode.bSetAuto:=FALSE; 
ELSIF stMode.iActMode=eAutoMode 
AND stMode.bSetSemi THEN; 
	stMode.bSetSemi:=FALSE;	
	stMode.iActMode:=eSemiAutoMode;
END_IF

IF stOperation.bStopResetAll THEN;
	stMode.bSetManual:=TRUE;
END_IF
END_ACTION

ACTION act_Reject_CMD:

	IF stMode.bSetManual 	THEN; sActErrorID:='300';END_IF	(*	'050x000x300',	'Warning',	'Manual mode request rejected, first pause automation',	*)
	IF stMode.bSetSemi 		THEN; sActErrorID:='301';END_IF	(*	'050x000x301',	'Warning',	'Semi mode request rejected, first pause automation',	*)
	IF stMode.bSetAuto 		THEN; sActErrorID:='302';END_IF	(*	'050x000x302',	'Warning',	'Auto mode request rejected, first pause automation',	*)
	act_GetErrorID_Format();
	fbPrintErrMessageByID(sFB_ModuleDescription:=sModuleDescription,sActErrorID:=sFullErrorId,bSFCError:=TRUE);
END_ACTION

ACTION act_SwitchFailed:

IF stMode.bSetManual 	THEN; sActErrorID:='303';END_IF	(*	'050x000x303',	'Warning',	'Manual mode request rejected, Pistion not in last auto pisition',	*)
IF stMode.bSetSemi 		THEN; sActErrorID:='304';END_IF	(*	'050x000x304',	'Warning',	'Semi mode request rejected, Pistion not in last auto pisition',	*)
IF stMode.bSetAuto 		THEN; sActErrorID:='304';END_IF	(*	'050x000x305',	'Warning',	'Auto mode request rejected, Pistion not in last auto pisition',	*)
act_GetErrorID_Format();
fbPrintErrMessageByID(sFB_ModuleDescription:=sModuleDescription,sActErrorID:=sFullErrorId,bSFCError:=TRUE);

stMode.bSetManual:=FALSE;
stMode.bSetSemi:=FALSE;
stMode.bSetAuto:=FALSE;
END_ACTION

ACTION Condition_Check_active:
bPistonsOK:=TRUE;
IF bPistonCheck THEN
	FOR i:=1 TO C_Max_Pistons DO;
		IF stPis[i].b_Exist
		AND (NOT stPis[i].st_SyncAuto) THEN;
			IF stPis[i].eModeZone=eModeZone THEN;
				stPis[i].b_Print_NotSyncAutoMessage:=TRUE;
				bPistonsOK:=FALSE;
			END_IF
		END_IF
	END_FOR	
END_IF
END_ACTION

ACTION Condition_Check_exit:
IF NOT bPistonsOK THEN;	
(*	IF stMode.bSetManual 	THEN; sActErrorID:='303';END_IF	(*	'050x000x303',	'Warning',	'Manual mode request rejected, Pistion not in last auto pisition',	*)
	IF stMode.bSetSemi 		THEN; sActErrorID:='304';END_IF	(*	'050x000x304',	'Warning',	'Semi mode request rejected, Pistion not in last auto pisition',	*)
	IF stMode.bSetAuto 		THEN; sActErrorID:='304';END_IF	(*	'050x000x305',	'Warning',	'Auto mode request rejected, Pistion not in last auto pisition',	*)
	act_GetErrorID_Format();
	fbPrintErrMessageByID(sModuleDescription:=sModuleDescription,sActErrorID:=sFullErrorId);*)
END_IF
END_ACTION

METHOD m_Error_zone_check : BOOL
VAR_INPUT
END_VAR

VAR
	i: INT;
	sCheckZone: STRING;

END_VAR
sCheckZone:=TO_STRING(stMode.eModeZone);

FOR i:=1 TO C_Max_Buffer_Act_list DO;
	IF TRUE 
	AND Buffer_Act_Message[i].sLevel='Error'
	AND Buffer_Act_Message[i].sModuleDescription=sCheckZone
	AND stOperation.iActOperation=E_OperationButtons.ePlayAll 
	THEN;
		stOperation.bSetPause:=TRUE;
	END_IF
END_FOR
END_METHOD

ACTION Ready_exit:
stOperation.bSetPause:=TRUE;
stOperation.iPauseHistory:=6;
END_ACTION

ACTION SetAuto_entry:
stMode.iActMode:=eAutoMode;
END_ACTION

ACTION SetMan_entry:
stMode.iActMode:=eManualMode;
END_ACTION

ACTION SetSemi_entry:
stMode.iActMode:=eSemiAutoMode;
END_ACTION

ACTION SwitchFail1_entry:
//entrance condition <NOT prg_Initialise.bGeneralDone>

//IF stMode.bSetAuto 		THEN; sActErrorID:='304';END_IF	(*	'050x000x305',	'Warning',	'Auto mode request rejected, Pistion not in last auto pisition',	*)

sActErrorID:='350'; // '050x000x350',	'Warning',	'Semi/Auto mode request rejected, initialize all system first',
act_GetErrorID_Format();
fbPrintErrMessageByID(sFB_ModuleDescription:=sModuleDescription,sActErrorID:=sFullErrorId,bSFCError:=TRUE);

stMode.bSetManual:=FALSE;
stMode.bSetSemi:=FALSE;
stMode.bSetAuto:=FALSE;
END_ACTION

END_FUNCTION_BLOCK

// ---- 00 Library/04-Messages/FB_PrintErrMessageByID_SFC_Cycle.TcPOU
FUNCTION_BLOCK FB_PrintErrMessageByID_SFC_Cycle
VAR_INPUT
	sActErrorID				: STRING;
	iFB_Num					: INT:=0;
	sFB_ModuleDescription	: STRING:='';
	bSFCError				: BOOL;
	sLast_ErrorToPrint		: STRING;
END_VAR
VAR_OUTPUT
END_VAR
VAR
	cFound				: INT;
	i					: INT;
	iFound				: INT;
	bNewMeasege			: BOOL;
	rtrig1				: R_TRIG;
	sLastErrorID		: STRING;
	sLastErrorID_ToPrint		: STRING;	
	j: INT;
	sActErrorID_List: STRING(11);
	sTemp1: STRING(11);
	sTemp2: STRING(11);
END_VAR


sLastErrorID_ToPrint:='';
	
IF bSFCError THEN
	IF sActErrorID<>'000x000x000'  AND sActErrorID<>'' THEN
		sLastErrorID:=sActErrorID;
		bNewMeasege:=TRUE;
		FOR i:=1 TO 100 DO
			IF Buffer_Act_Message[i].sErrID=sActErrorID THEN;
				//IF Buffer_Act_Message[i].sModuleDescription = sFB_ModuleDescription THEN
					bNewMeasege:=FALSE;
					EXIT; 
				//END_IF
			END_IF
		END_FOR
	ELSE
		bNewMeasege:=FALSE;
	END_IF
	
	
	IF bNewMeasege THEN;
		FOR i:=100 TO 2 BY -1 DO
			Buffer_Act_Message[i].sDateTime:=Buffer_Act_Message[i-1].sDateTime;
			Buffer_Act_Message[i].sErrID:=Buffer_Act_Message[i-1].sErrID;
			Buffer_Act_Message[i].sErrorMessage:=Buffer_Act_Message[i-1].sErrorMessage;
			Buffer_Act_Message[i].sLevel:=Buffer_Act_Message[i-1].sLevel;
			Buffer_Act_Message[i].sModuleDescription:=Buffer_Act_Message[i-1].sModuleDescription;
		END_FOR
		
		Buffer_Act_Message[1].sDateTime:=prg_RealClock.sRealTime_Date;
		Buffer_Act_Message[1].sErrID:=sActErrorID;
		Buffer_Act_Message[1].sModuleDescription:=sFB_ModuleDescription;

		IF REPLACE(sActErrorID,'',8,1)='PUZ' THEN;
			sActErrorID_List:=REPLACE(sActErrorID,'000x000',7,1);	
			sTemp1:=sActErrorID_List;		
		ELSE;
			sActErrorID_List:=REPLACE(sActErrorID,'000',3,5);
			sTemp2:=sActErrorID_List;
		END_IF
		
		
		IF sActErrorID='000x000x999' THEN;
			Buffer_Act_Message[1].sErrorMessage:=CONCAT('Cycle message: ',sLast_ErrorToPrint);
			Buffer_Act_Message[1].sLevel:='Error';
		ELSE
			cFound:=0;
			FOR i:=1 TO C_Max_ErrorList DO
				IF ar_ErrorList[i,eErrID]=sActErrorID_List THEN
					iFound:=i;
					ar_ErrorActive[iFound]:=TRUE;
					cFound:=cFound+1;
				END_IF
			END_FOR
	
			IF cFound=1 THEN;
				Buffer_Act_Message[1].sErrorMessage:=ar_ErrorList[iFound,eErrMeassage];	(*	Error from the List	*)
				Buffer_Act_Message[1].sLevel:=ar_ErrorList[iFound,eErrLevel];	(*	Error Level from the List	*)
			ELSIF cFound=0 THEN; //(*	Error ID not Foud on the List	*)
				//Buffer_Act_Message[1].sErrorMessage:='Error ID not found on the "Error_List"';
				Buffer_Act_Message[1].sErrorMessage:=CONCAT('Cycle message[1]: ',sLast_ErrorToPrint);
				Buffer_Act_Message[1].sLevel:='Error';
			ELSIF cFound>1 THEN; //(*	More then one Errors Foud with the same  ID		*)
				//Buffer_Act_Message[1].sErrorMessage:='More then one error with the same ID  found on the "Error_list"';
				Buffer_Act_Message[1].sErrorMessage:=CONCAT('Cycle message[2]: ',sLast_ErrorToPrint);
				Buffer_Act_Message[1].sLevel:='Error';
			END_IF
		END_IF
		FUN_Write_Line_To_History();
	END_IF
	
END_IF

(*
rtrig1(CLK:= NOT bSFCError , Q=> );
IF rtrig1.Q THEN  // if cycle not in pause
	FOR i:= 2 TO 100 DO //loop for search 
		IF Buffer_Act_Message[i-1].sErrID = sLastErrorID THEN // search if last error id = buffer which it error table.
			FOR j:= i TO 100 DO //if found message id then delete it.
				Buffer_Act_Message[j-1]:=Buffer_Act_Message[j];//delete
			END_FOR
		END_IF
	END_FOR
END_IF
*)

END_FUNCTION_BLOCK

// ---- 00 Library/07-Mode/FB_Operation.TcPOU
FUNCTION_BLOCK FB_Operation
VAR_INPUT
	bStateSafe: BOOL:=TRUE;
END_VAR
VAR
	r1: R_TRIG;
	r2: R_TRIG;
	arPauseHistory: ARRAY[0..9] OF INT;
	ton_StopResetAllTime: TON;
	ton_PauseDelay: TON;
END_VAR
VAR_IN_OUT
	stOper	:ST_OperationButtons;
END_VAR

r1(CLK:=stOper.bSetPlay,Q=>stOper.b_rt_Play );
IF  r1.Q THEN
	stOper.iActOperation:=E_OperationButtons.ePlayAll;
	stOper.bSetPause:=FALSE;
	stOper.bSetPlay:=FALSE;
END_IF

IF stOper.bSetPlay OR stOper.iActOperation=E_OperationButtons.ePlayAll THEN;
	stOper.bSetPlay:=FALSE;
END_IF

r2(CLK:= stOper.bSetPause, Q=>stOper.b_rt_Pause );
IF r2.Q THEN
	stOper.iActOperation:=E_OperationButtons.ePauseAll;
	stOper.bSetPause:=FALSE;
	stOper.bSetPlay:=FALSE;
	m_WritePauseHystory(iVar:=stOper.iPauseHistory);
END_IF

IF stOper.bSetPause OR stOper.iActOperation=E_OperationButtons.ePauseAll THEN;
	stOper.bSetPause:=FALSE;
END_IF

ton_StopResetAllTime(PT:=T#0.5S);
IF stOper.bStopResetAll OR NOT bStateSafe THEN;
	ton_StopResetAllTime.IN:=TRUE;
	stOper.bStopResetAll:=TRUE;
	IF ton_StopResetAllTime.Q THEN;
		ton_StopResetAllTime.IN:=FALSE;
		stOper.bStopResetAll:=FALSE;
	END_IF
END_IF

ton_PauseDelay(PT:=T#2S,
IN:=stOper.iActOperation=E_OperationButtons.ePauseAll,
Q=>stOper.bPauseOnDelayed
);

METHOD m_WritePauseHystory : BOOL
VAR_IN_OUT
	iVar: INT;

END_VAR
VAR
	i: INT;
END_VAR
FOR i:=9 TO 1 BY -1 DO;
	arPauseHistory[i]:=arPauseHistory[i-1];
END_FOR
arPauseHistory[0]:=iVar;
iVar:=0;
END_METHOD

END_FUNCTION_BLOCK

// ---- 01 Instance/07-Mode/prg_LightTower.TcPOU
PROGRAM prg_LightTower
VAR_INPUT
	bBuzzerBypass: BOOL;
END_VAR
VAR

	ton_Blink				: TON;
	ton_Buzzer				: TON;
	t_Buzzer				: TIME:=T#2S;
	t_BuzzerShort			: TIME:=T#0.5S;
	t_BuzzerErrorDelay		: TIME:=T#10S;
	t_BuzzerWarningDelay	: TIME:=T#30S;
	//eLightTowerState_Last	: E_LightTowerState;
	bBuzzerMuteMemo: BOOL;	
	ton_MuteBuzzer: TON;
	ton_NoMessage: TON;
	ton_BuzzerLongTimeOn: TON;
END_VAR

VAR_OUTPUT
	qLedGreen	: BOOL;
	qLedYellow	: BOOL;
	qLedRed		: BOOL;
	qBuzzer		: BOOL;	
END_VAR

// Interface
(*
q_EL[1].ch1:=qLedGreen;
q_EL[1].ch2:=qLedYellow;
q_EL[1].ch3:=qLedRed;
q_EL[1].ch4:=qBuzzer;
*)
//.....................
(*
TYPE E_LightTowerState :
(
	eLightsOff := 0,
	eRed,				//Error
	eYellow,			//Pause
	eGreen,				//Run
	eGreenYellowBlink	//Run and warning
);
END_TYPE
*)
act_Operation();
ton_Blink(IN:=NOT ton_Blink.Q);
CASE eLightTowerState OF
	eLightsOff:;
		qLedGreen	:=FALSE;
		qLedYellow	:=FALSE;
		qLedRed		:=FALSE;
		eBuzzerMode:=eBuzzerOff;	
		
	eGreen:;
		qLedGreen	:=TRUE;
		qLedYellow	:=FALSE;
		qLedRed		:=FALSE;
		eBuzzerMode:=eBuzzerOff;	
		
	eGreen_YellowBlink:;
		qLedGreen	:=TRUE;
		qLedYellow	:=TRUE;
		qLedRed		:=FALSE;
		IF bBuzzerMuteMemo THEN;
			eBuzzerMode:=eBuzzerOff;
		ELSE
			eBuzzerMode:=eBuzzerWarning;
		END_IF
		ton_Blink.PT:=T#1S;
		IF ton_Blink.ET>T#0.5S THEN; qLedYellow:=FALSE; ELSE;qLedGreen:=FALSE; END_IF	
		
	eGreenBlink:;
		qLedGreen	:=TRUE;
		qLedYellow	:=FALSE;
		qLedRed		:=FALSE;
		eBuzzerMode:=eBuzzerOff;		
		ton_Blink.PT:=T#1S;
		IF ton_Blink.ET>T#0.5S THEN; qLedGreen:=FALSE; END_IF	

	eGreenBlink_YellowBlink:;
		qLedGreen	:=TRUE;
		qLedYellow	:=TRUE;
		qLedRed		:=FALSE;
		IF bBuzzerMuteMemo THEN;
			eBuzzerMode:=eBuzzerOff;
		ELSE
			eBuzzerMode:=eBuzzerWarning;
		END_IF
		ton_Blink.PT:=T#1S;
		IF ton_Blink.ET>T#0.5S THEN; qLedYellow:=FALSE; ELSE;qLedGreen:=FALSE; END_IF

	eGreenBlink_RedBlink:;
		qLedGreen	:=TRUE;
		qLedYellow	:=FALSE;
		qLedRed		:=TRUE;
		IF bBuzzerMuteMemo THEN;
			eBuzzerMode:=eBuzzerOff;
		ELSE
			eBuzzerMode:=eBuzzerError;
		END_IF
		ton_Blink.PT:=T#1S;
		IF ton_Blink.ET>T#0.5S THEN; qLedRed:=FALSE; ELSE;qLedGreen:=FALSE; END_IF
		
	eYellow:;
		qLedGreen	:=FALSE;
		qLedYellow	:=TRUE;
		qLedRed		:=FALSE;
		eBuzzerMode:=eBuzzerOff;	
		
	eRed:;
		qLedGreen	:=FALSE;
		qLedYellow	:=FALSE;
		qLedRed		:=TRUE;
		IF bBuzzerMuteMemo THEN;
			eBuzzerMode:=eBuzzerOff;
		ELSE
			eBuzzerMode:=eBuzzerError;
		END_IF
END_CASE

ton_NoMessage(PT:=T#5S,IN:=bBuzzerMuteMemo AND iActErrors=0 AND iActWarning=0);

IF (stOpMain.bSetPlay
	(*OR stOpLoad.bSetPlay
	OR stOpUnload.bSetPlay
	OR stOpManip.bSetPlay
	OR stOpHMI.bSetPlay
	OR prg_Call_OpMode.fbModeIndex.rt_Play.Q
	OR prg_Call_OpMode.fbModeLoad.rt_Play.Q
	OR prg_Call_OpMode.fbModeUnload.rt_Play.Q
	OR prg_Call_OpMode.fbModeManip.rt_Play.Q*)
	OR ton_NoMessage.Q	
)
THEN;
	ton_MuteBuzzer.IN:=TRUE;
END_IF
IF ton_MuteBuzzer.IN THEN;
	bBuzzerMuteMemo:=FALSE;
END_IF
ton_MuteBuzzer(PT:=T#1S);
IF ton_MuteBuzzer.Q THEN
	ton_MuteBuzzer.IN:=FALSE;
END_IF
IF prg_Messages.ResetErrors OR ton_BuzzerLongTimeOn.Q THEN;// iActErrors=0 AND iActWarning=0
	bBuzzerMuteMemo:=TRUE;
END_IF
ton_BuzzerLongTimeOn(PT:=T#30M,IN:=eBuzzerMode<>eBuzzerOff);

(*
TYPE E_BuzzerMode :
(
	eBuzzerOff := 0,
	eBuzzerError,		//Short Delay Off
	eBuzzerWarning		//Long Delay Off
);
END_TYPE
*)

IF NOT bBuzzerBypass THEN
	ton_Buzzer();
	CASE eBuzzerMode OF
		eBuzzerOff :;
			qBuzzer:=FALSE;
			
			ton_Buzzer.IN:=FALSE;
		eBuzzerError:;			//Short Delay Off
			qBuzzer:=TRUE;
			ton_Buzzer.PT:=t_BuzzerErrorDelay;
			ton_Buzzer.IN:=NOT ton_Buzzer.Q;
			IF ton_Buzzer.ET>t_Buzzer THEN; qBuzzer:=FALSE; END_IF
		eBuzzerWarning:;		//Long Delay Off
			qBuzzer:=TRUE;
			ton_Buzzer.PT:=t_BuzzerWarningDelay;
			ton_Buzzer.IN:=NOT ton_Buzzer.Q;
			IF ton_Buzzer.ET>t_BuzzerShort THEN; qBuzzer:=FALSE; END_IF
	END_CASE	
ELSE
	qBuzzer:=FALSE;
END_IF

ACTION act_Operation:
IF 		stOpMain.iActOperation=E_OperationButtons.ePauseAll
	AND iActErrors<>0
	THEN;	
	eLightTowerState:=E_LightTowerState.eRed;
 						//7
ELSIF 	stOpMain.iActOperation=E_OperationButtons.ePauseAll
	AND iActErrors=0
	THEN;
	eLightTowerState:=E_LightTowerState.eYellow;					//6	
	
ELSIF 	stOpMain.iActOperation=E_OperationButtons.ePlayAll
	AND iActErrors=0
 	AND iActWarning<>0
	THEN;
	eLightTowerState:=E_LightTowerState.eGreenBlink_YellowBlink;	//4
		
ELSIF 	stOpMain.iActOperation=E_OperationButtons.ePlayAll
	AND iActErrors=0 
	AND iActWarning=0 
	THEN;
	eLightTowerState:=E_LightTowerState.eGreen;						//1
END_IF
END_ACTION

ACTION act_Operation_Multi:
IF 		stOpMain.iActOperation=E_OperationButtons.ePauseAll
	//AND stOpLoad.iActOperation=E_OperationButtons.ePauseAll
	//AND stOpUnload.iActOperation=E_OperationButtons.ePauseAll
	//AND stOpManip.iActOperation=E_OperationButtons.ePauseAll
	//AND stOpHMI.iActOperation=E_OperationButtons.ePauseAll
	AND iActErrors<>0
	THEN;	
	eLightTowerState:=E_LightTowerState.eRed;
 						//7
ELSIF 	stOpMain.iActOperation=E_OperationButtons.ePauseAll
	//AND stOpLoad.iActOperation=E_OperationButtons.ePauseAll
	//AND stOpUnload.iActOperation=E_OperationButtons.ePauseAll
	//AND stOpManip.iActOperation=E_OperationButtons.ePauseAll
	//AND stOpHMI.iActOperation=E_OperationButtons.ePauseAll
	AND iActErrors=0
	THEN;
	eLightTowerState:=E_LightTowerState.eYellow;					//6
	
ELSIF 	(stOpMain.iActOperation=E_OperationButtons.ePlayAll
	(*OR stOpLoad.iActOperation=E_OperationButtons.ePlayAll
	OR stOpUnload.iActOperation=E_OperationButtons.ePlayAll
	OR stOpManip.iActOperation=E_OperationButtons.ePlayAll
	OR stOpHMI.iActOperation=E_OperationButtons.ePlayAll*))
	AND iActErrors<>0 
	THEN;
	eLightTowerState:=E_LightTowerState.eGreenBlink_RedBlink;		//5
	
ELSIF 	(stOpMain.iActOperation=E_OperationButtons.ePlayAll
	(*OR stOpLoad.iActOperation=E_OperationButtons.ePlayAll
	OR stOpUnload.iActOperation=E_OperationButtons.ePlayAll
	OR stOpManip.iActOperation=E_OperationButtons.ePlayAll
	OR stOpHMI.iActOperation=E_OperationButtons.ePlayAll*))
	AND iActErrors=0
 	AND iActWarning<>0
	THEN;
	eLightTowerState:=E_LightTowerState.eGreenBlink_YellowBlink;	//4
	
ELSIF  	(stOpMain.iActOperation=E_OperationButtons.ePlayAll
	(*OR stOpLoad.iActOperation=E_OperationButtons.ePlayAll
	OR stOpUnload.iActOperation=E_OperationButtons.ePlayAll
	OR stOpManip.iActOperation=E_OperationButtons.ePlayAll
	OR stOpHMI.iActOperation=E_OperationButtons.ePlayAll*))
	AND  (stOpMain.iActOperation=E_OperationButtons.ePauseAll
	(*OR stOpLoad.iActOperation=E_OperationButtons.ePauseAll
	OR stOpUnload.iActOperation=E_OperationButtons.ePauseAll
	OR stOpManip.iActOperation=E_OperationButtons.ePauseAll
	OR stOpHMI.iActOperation=E_OperationButtons.ePauseAll*))	
	AND iActErrors=0
 	AND iActWarning=0
	THEN;
	eLightTowerState:=E_LightTowerState.eGreenBlink;				//3
	
ELSIF 	stOpMain.iActOperation=E_OperationButtons.ePlayAll
	(*AND stOpLoad.iActOperation=E_OperationButtons.ePlayAll
	AND stOpUnload.iActOperation=E_OperationButtons.ePlayAll
	AND stOpManip.iActOperation=E_OperationButtons.ePlayAll
	AND stOpHMI.iActOperation=E_OperationButtons.ePlayAll*)
	AND iActErrors=0 
	AND iActWarning<>0
	THEN;
	eLightTowerState:=E_LightTowerState.eGreen_YellowBlink;			//2
	
ELSIF 	stOpMain.iActOperation=E_OperationButtons.ePlayAll
	(*AND stOpLoad.iActOperation=E_OperationButtons.ePlayAll
	AND stOpUnload.iActOperation=E_OperationButtons.ePlayAll
	AND stOpManip.iActOperation=E_OperationButtons.ePlayAll
	AND stOpHMI.iActOperation=E_OperationButtons.ePlayAll*)
	AND iActErrors=0 
	AND iActWarning=0 
	THEN;
	eLightTowerState:=E_LightTowerState.eGreen;						//1
END_IF
END_ACTION

END_PROGRAM

// ---- 01 Instance/07-Mode/FB_LightTower.TcPOU
FUNCTION_BLOCK FB_LightTower
VAR_INPUT
	bBuzzerBypass: BOOL;
END_VAR
VAR_OUTPUT
	qLedGreen	: BOOL;
	qLedYellow	: BOOL;
	qLedRed		: BOOL;
	qLedBlue	: BOOL;
	qBuzzer		: BOOL;		
	
	qSignal_1: BOOL; //wire BN
	qSignal_2: BOOL; //wire GY
	qSignal_3: BOOL; //wire BK
	qSignal_4: BOOL; //wire WT

END_VAR
VAR
	eLightTowerState		: E_LightTowerState;
	eLightTower_Type		: E_LightTower_Type:=E_LightTower_Type.eSingleLayer;

	
	ton_Blink				: TON;
	ton_Buzzer				: TON;
	t_Buzzer				: TIME:=T#2S;
	t_BuzzerShort			: TIME:=T#0.5S;
	t_BuzzerErrorDelay		: TIME:=T#10S;
	t_BuzzerWarningDelay	: TIME:=T#30S;
	//eLightTowerState_Last	: E_LightTowerState;
	bBuzzerMuteMemo: BOOL;	
	ton_MuteBuzzer: TON;
	ton_NoMessage: TON;
	ton_BuzzerLongTimeOn: TON;	
END_VAR

ton_Blink(IN:=NOT ton_Blink.Q);
CASE eLightTower_Type OF
	E_LightTower_Type.eSingleLayer: m_Single_Layer();
	E_LightTower_Type.eMultiLayer: m_Multi_Layer();
	
END_CASE


ton_NoMessage(PT:=T#5S,IN:=bBuzzerMuteMemo AND iActErrors=0 AND iActWarning=0);

IF (stOpMain.bSetPlay
	(*OR stOpLoad.bSetPlay
	OR stOpUnload.bSetPlay
	OR stOpManip.bSetPlay
	OR stOpHMI.bSetPlay
	OR prg_Call_OpMode.fbModeIndex.rt_Play.Q
	OR prg_Call_OpMode.fbModeLoad.rt_Play.Q
	OR prg_Call_OpMode.fbModeUnload.rt_Play.Q
	OR prg_Call_OpMode.fbModeManip.rt_Play.Q*)
	OR ton_NoMessage.Q	
)
THEN;
	ton_MuteBuzzer.IN:=TRUE;
END_IF
IF ton_MuteBuzzer.IN THEN;
	bBuzzerMuteMemo:=FALSE;
END_IF
ton_MuteBuzzer(PT:=T#1S);
IF ton_MuteBuzzer.Q THEN
	ton_MuteBuzzer.IN:=FALSE;
END_IF
IF prg_Messages.ResetErrors OR ton_BuzzerLongTimeOn.Q THEN;// iActErrors=0 AND iActWarning=0
	bBuzzerMuteMemo:=TRUE;
END_IF
ton_BuzzerLongTimeOn(PT:=T#30M,IN:=eBuzzerMode<>eBuzzerOff);

(*
TYPE E_BuzzerMode :
(
	eBuzzerOff := 0,
	eBuzzerError,		//Short Delay Off
	eBuzzerWarning		//Long Delay Off
);
END_TYPE
*)

IF NOT bBuzzerBypass THEN
	ton_Buzzer();
	CASE eBuzzerMode OF
		eBuzzerOff :;
			qBuzzer:=FALSE;
			
			ton_Buzzer.IN:=FALSE;
		eBuzzerError:;			//Short Delay Off
			qBuzzer:=TRUE;
			ton_Buzzer.PT:=t_BuzzerErrorDelay;
			ton_Buzzer.IN:=NOT ton_Buzzer.Q;
			IF ton_Buzzer.ET>t_Buzzer THEN; qBuzzer:=FALSE; END_IF
		eBuzzerWarning:;		//Long Delay Off
			qBuzzer:=TRUE;
			ton_Buzzer.PT:=t_BuzzerWarningDelay;
			ton_Buzzer.IN:=NOT ton_Buzzer.Q;
			IF ton_Buzzer.ET>t_BuzzerShort THEN; qBuzzer:=FALSE; END_IF
	END_CASE	
ELSE
	qBuzzer:=FALSE;
END_IF

METHOD m_Multi_Layer : BOOL
VAR_INPUT
END_VAR
CASE eLightTowerState OF
	E_LightTowerState.eLightsOff:;
		qLedGreen	:=FALSE;
		qLedYellow	:=FALSE;
		qLedRed		:=FALSE;
		qLedBlue	:=FALSE;
		eBuzzerMode:=eBuzzerOff;	
		
	E_LightTowerState.eGreen:;
		qLedGreen	:=TRUE;
		qLedYellow	:=FALSE;
		qLedRed		:=FALSE;
		qLedBlue	:=FALSE;
		eBuzzerMode:=eBuzzerOff;	
		
	E_LightTowerState.eGreen_YellowBlink:;
		qLedGreen	:=TRUE;
		qLedYellow	:=TRUE;
		qLedRed		:=FALSE;
		qLedBlue	:=FALSE;
		IF bBuzzerMuteMemo THEN;
			eBuzzerMode:=eBuzzerOff;
		ELSE
			eBuzzerMode:=eBuzzerWarning;
		END_IF
		ton_Blink.PT:=T#1S;
		IF ton_Blink.ET>T#0.5S THEN; qLedYellow:=FALSE; ELSE;qLedGreen:=FALSE; END_IF	
		
	E_LightTowerState.eGreenBlink:;
		qLedGreen	:=TRUE;
		qLedYellow	:=FALSE;
		qLedRed		:=FALSE;
		qLedBlue	:=FALSE;
		eBuzzerMode:=eBuzzerOff;		
		ton_Blink.PT:=T#1S;
		IF ton_Blink.ET>T#0.5S THEN; qLedGreen:=FALSE; END_IF	

	E_LightTowerState.eGreenBlink_YellowBlink:;
		qLedGreen	:=TRUE;
		qLedYellow	:=TRUE;
		qLedRed		:=FALSE;
		qLedBlue	:=FALSE;
		IF bBuzzerMuteMemo THEN;
			eBuzzerMode:=eBuzzerOff;
		ELSE
			eBuzzerMode:=eBuzzerWarning;
		END_IF
		ton_Blink.PT:=T#1S;
		IF ton_Blink.ET>T#0.5S THEN; qLedYellow:=FALSE; ELSE;qLedGreen:=FALSE; END_IF

	E_LightTowerState.eGreenBlink_RedBlink:;
		qLedGreen	:=TRUE;
		qLedYellow	:=FALSE;
		qLedRed		:=TRUE;
		qLedBlue	:=FALSE;
		IF bBuzzerMuteMemo THEN;
			eBuzzerMode:=eBuzzerOff;
		ELSE
			eBuzzerMode:=eBuzzerError;
		END_IF
		ton_Blink.PT:=T#1S;
		IF ton_Blink.ET>T#0.5S THEN; qLedRed:=FALSE; ELSE;qLedGreen:=FALSE; END_IF
		
	E_LightTowerState.eYellow:;
		qLedGreen	:=FALSE;
		qLedYellow	:=TRUE;
		qLedRed		:=FALSE;
		qLedBlue	:=FALSE;
		eBuzzerMode:=eBuzzerOff;	
		
	E_LightTowerState.eRed:;
		qLedGreen	:=FALSE;
		qLedYellow	:=FALSE;
		qLedRed		:=TRUE;
		qLedBlue	:=FALSE;
		IF bBuzzerMuteMemo THEN;
			eBuzzerMode:=eBuzzerOff;
		ELSE
			eBuzzerMode:=eBuzzerError;
		END_IF
		
	E_LightTowerState.eBlue:;
		qLedGreen	:=FALSE;
		qLedYellow	:=FALSE;
		qLedRed		:=FALSE;
		qLedBlue	:=TRUE;
		eBuzzerMode:=eBuzzerOff;	
				
END_CASE
END_METHOD

METHOD m_Op_Case1 : BOOL
VAR_INPUT
END_VAR
IF 		stOpMain.iActOperation=E_OperationButtons.ePauseAll
	AND iActErrors<>0
	THEN;	
	eLightTowerState:=E_LightTowerState.eRed;
 						//7
ELSIF 	stOpMain.iActOperation=E_OperationButtons.ePauseAll
	AND iActErrors=0
	THEN;
	eLightTowerState:=E_LightTowerState.eYellow;					//6	
	
ELSIF 	stOpMain.iActOperation=E_OperationButtons.ePlayAll
	AND iActErrors=0
 	AND iActWarning<>0
	THEN;
	eLightTowerState:=E_LightTowerState.eGreenBlink_YellowBlink;	//4
		
ELSIF 	stOpMain.iActOperation=E_OperationButtons.ePlayAll
	AND iActErrors=0 
	AND iActWarning=0 
	THEN;
	eLightTowerState:=E_LightTowerState.eGreen;						//1
END_IF
END_METHOD

METHOD m_Op_Case2 : BOOL
VAR_INPUT
END_VAR
IF 		stOpMain.iActOperation=E_OperationButtons.ePauseAll
	//AND stOpLoad.iActOperation=E_OperationButtons.ePauseAll
	//AND stOpUnload.iActOperation=E_OperationButtons.ePauseAll
	//AND stOpManip.iActOperation=E_OperationButtons.ePauseAll
	//AND stOpHMI.iActOperation=E_OperationButtons.ePauseAll
	AND iActErrors<>0
	THEN;	
	eLightTowerState:=E_LightTowerState.eRed;
 						//7
ELSIF 	stOpMain.iActOperation=E_OperationButtons.ePauseAll
	//AND stOpLoad.iActOperation=E_OperationButtons.ePauseAll
	//AND stOpUnload.iActOperation=E_OperationButtons.ePauseAll
	//AND stOpManip.iActOperation=E_OperationButtons.ePauseAll
	//AND stOpHMI.iActOperation=E_OperationButtons.ePauseAll
	AND iActErrors=0
	THEN;
	eLightTowerState:=E_LightTowerState.eYellow;					//6
	
ELSIF 	(stOpMain.iActOperation=E_OperationButtons.ePlayAll
	(*OR stOpLoad.iActOperation=E_OperationButtons.ePlayAll
	OR stOpUnload.iActOperation=E_OperationButtons.ePlayAll
	OR stOpManip.iActOperation=E_OperationButtons.ePlayAll
	OR stOpHMI.iActOperation=E_OperationButtons.ePlayAll*))
	AND iActErrors<>0 
	THEN;
	eLightTowerState:=E_LightTowerState.eGreenBlink_RedBlink;		//5
	
ELSIF 	(stOpMain.iActOperation=E_OperationButtons.ePlayAll
	(*OR stOpLoad.iActOperation=E_OperationButtons.ePlayAll
	OR stOpUnload.iActOperation=E_OperationButtons.ePlayAll
	OR stOpManip.iActOperation=E_OperationButtons.ePlayAll
	OR stOpHMI.iActOperation=E_OperationButtons.ePlayAll*))
	AND iActErrors=0
 	AND iActWarning<>0
	THEN;
	eLightTowerState:=E_LightTowerState.eGreenBlink_YellowBlink;	//4
	
ELSIF  	(stOpMain.iActOperation=E_OperationButtons.ePlayAll
	(*OR stOpLoad.iActOperation=E_OperationButtons.ePlayAll
	OR stOpUnload.iActOperation=E_OperationButtons.ePlayAll
	OR stOpManip.iActOperation=E_OperationButtons.ePlayAll
	OR stOpHMI.iActOperation=E_OperationButtons.ePlayAll*))
	AND  (stOpMain.iActOperation=E_OperationButtons.ePauseAll
	(*OR stOpLoad.iActOperation=E_OperationButtons.ePauseAll
	OR stOpUnload.iActOperation=E_OperationButtons.ePauseAll
	OR stOpManip.iActOperation=E_OperationButtons.ePauseAll
	OR stOpHMI.iActOperation=E_OperationButtons.ePauseAll*))	
	AND iActErrors=0
 	AND iActWarning=0
	THEN;
	eLightTowerState:=E_LightTowerState.eGreenBlink;				//3
	
ELSIF 	stOpMain.iActOperation=E_OperationButtons.ePlayAll
	(*AND stOpLoad.iActOperation=E_OperationButtons.ePlayAll
	AND stOpUnload.iActOperation=E_OperationButtons.ePlayAll
	AND stOpManip.iActOperation=E_OperationButtons.ePlayAll
	AND stOpHMI.iActOperation=E_OperationButtons.ePlayAll*)
	AND iActErrors=0 
	AND iActWarning<>0
	THEN;
	eLightTowerState:=E_LightTowerState.eGreen_YellowBlink;			//2
	
ELSIF 	stOpMain.iActOperation=E_OperationButtons.ePlayAll
	(*AND stOpLoad.iActOperation=E_OperationButtons.ePlayAll
	AND stOpUnload.iActOperation=E_OperationButtons.ePlayAll
	AND stOpManip.iActOperation=E_OperationButtons.ePlayAll
	AND stOpHMI.iActOperation=E_OperationButtons.ePlayAll*)
	AND iActErrors=0 
	AND iActWarning=0 
	THEN;
	eLightTowerState:=E_LightTowerState.eGreen;						//1
END_IF
END_METHOD

METHOD m_Op_Case3 : BOOL
VAR_INPUT
END_VAR
END_METHOD

METHOD m_Single_Layer : BOOL
VAR_INPUT
END_VAR
CASE eLightTowerState OF
	E_LightTowerState.eLightsOff:;
		qLedGreen	:=FALSE;
		qLedYellow	:=FALSE;
		qLedRed		:=FALSE;
		qLedBlue	:=FALSE;
		eBuzzerMode:=eBuzzerOff;	
		
	E_LightTowerState.eGreen:;
		qLedGreen	:=TRUE;
		qLedYellow	:=FALSE;
		qLedRed		:=FALSE;
		qLedBlue	:=FALSE;
		eBuzzerMode:=eBuzzerOff;	
		
	E_LightTowerState.eGreen_YellowBlink:;
		qLedGreen	:=TRUE;
		qLedYellow	:=TRUE;
		qLedRed		:=FALSE;
		qLedBlue	:=FALSE;
		IF bBuzzerMuteMemo THEN;
			eBuzzerMode:=eBuzzerOff;
		ELSE
			eBuzzerMode:=eBuzzerWarning;
		END_IF
		ton_Blink.PT:=T#1S;
		IF ton_Blink.ET>T#0.5S THEN; qLedYellow:=FALSE; ELSE;qLedGreen:=FALSE; END_IF	
		
	E_LightTowerState.eGreenBlink:;
		qLedGreen	:=TRUE;
		qLedYellow	:=FALSE;
		qLedRed		:=FALSE;
		qLedBlue	:=FALSE;
		eBuzzerMode:=eBuzzerOff;		
		ton_Blink.PT:=T#1S;
		IF ton_Blink.ET>T#0.5S THEN; qLedGreen:=FALSE; END_IF	

	E_LightTowerState.eGreenBlink_YellowBlink:;
		qLedGreen	:=TRUE;
		qLedYellow	:=TRUE;
		qLedRed		:=FALSE;
		qLedBlue	:=FALSE;
		IF bBuzzerMuteMemo THEN;
			eBuzzerMode:=eBuzzerOff;
		ELSE
			eBuzzerMode:=eBuzzerWarning;
		END_IF
		ton_Blink.PT:=T#1S;
		IF ton_Blink.ET>T#0.5S THEN; qLedYellow:=FALSE; ELSE;qLedGreen:=FALSE; END_IF

	E_LightTowerState.eGreenBlink_RedBlink:;
		qLedGreen	:=TRUE;
		qLedYellow	:=FALSE;
		qLedRed		:=TRUE;
		qLedBlue	:=FALSE;
		IF bBuzzerMuteMemo THEN;
			eBuzzerMode:=eBuzzerOff;
		ELSE
			eBuzzerMode:=eBuzzerError;
		END_IF
		ton_Blink.PT:=T#1S;
		IF ton_Blink.ET>T#0.5S THEN; qLedRed:=FALSE; ELSE;qLedGreen:=FALSE; END_IF
		
	E_LightTowerState.eYellow:;
		qLedGreen	:=FALSE;
		qLedYellow	:=TRUE;
		qLedRed		:=FALSE;
		qLedBlue	:=FALSE;
		eBuzzerMode:=eBuzzerOff;	
		
	E_LightTowerState.eRed:;
		qLedGreen	:=FALSE;
		qLedYellow	:=FALSE;
		qLedRed		:=TRUE;
		qLedBlue	:=FALSE;
		IF bBuzzerMuteMemo THEN;
			eBuzzerMode:=eBuzzerOff;
		ELSE
			eBuzzerMode:=eBuzzerError;
		END_IF
		
	E_LightTowerState.eBlue:;
		qLedGreen	:=FALSE;
		qLedYellow	:=FALSE;
		qLedRed		:=FALSE;
		qLedBlue	:=TRUE;
		eBuzzerMode:=eBuzzerOff;	
				
END_CASE


IF qLedRed THEN;
	qSignal_1:=TRUE;	//wire BN
	qSignal_2:=FALSE;	//wire GY
	qSignal_3:=FALSE;	//wire BK
	qSignal_4:=FALSE;	//wire WT	
ELSIF qLedYellow THEN;
	qSignal_1:=TRUE;	//wire BN
	qSignal_2:=FALSE;	//wire GY
	qSignal_3:=FALSE;	//wire BK
	qSignal_4:=TRUE;	//wire WT	
ELSIF qLedGreen THEN;
	qSignal_1:=FALSE;	//wire BN
	qSignal_2:=FALSE;	//wire GY
	qSignal_3:=FALSE;	//wire BK
	qSignal_4:=TRUE;	//wire WT	
ELSIF qLedBlue THEN;
	qSignal_1:=FALSE;	//wire BN
	qSignal_2:=TRUE;	//wire GY
	qSignal_3:=FALSE;	//wire BK
	qSignal_4:=FALSE;	//wire WT	
ELSE;
	qSignal_1:=FALSE;	//wire BN
	qSignal_2:=FALSE;	//wire GY
	qSignal_3:=FALSE;	//wire BK
	qSignal_4:=FALSE;	//wire WT
END_IF
END_METHOD

PROPERTY pState : E_LightTowerState
GET
pState:=eLightTowerState;
END_GET
SET
eLightTowerState:=pState;
END_SET
END_PROPERTY

END_FUNCTION_BLOCK

// ---- 01 Instance/07-Mode/FB_LightTower_Control.TcPOU
FUNCTION_BLOCK FB_LightTower_Control
VAR_INPUT
	ES_State		: BOOL;
	RunProcess1		: BOOL;
	RunProcess2		: BOOL;
	RunProcess3		: BOOL;
	ModeZone1		: E_ModeZone;
	ModeZone2		: E_ModeZone;
	ModeZone3		: E_ModeZone;
END_VAR

VAR_OUTPUT
	eLightTowerState		: E_LightTowerState;
END_VAR
VAR
END_VAR

IF ES_State THEN;
	IF stOper[ModeZone1].iActOperation=E_OperationButtons.ePauseAll 
	OR stOper[ModeZone2].iActOperation=E_OperationButtons.ePauseAll
	OR stOper[ModeZone3].iActOperation=E_OperationButtons.ePauseAll
	THEN;
		eLightTowerState:= E_LightTowerState.eYellow;
	ELSIF RunProcess1 OR RunProcess2 OR RunProcess3 THEN;
		eLightTowerState:= E_LightTowerState.eGreen;
	ELSE;
		eLightTowerState:= E_LightTowerState.eBlue;
	END_IF
	
ELSE;
	eLightTowerState:= E_LightTowerState.eRed;
END_IF

END_FUNCTION_BLOCK

// ---- 00 Library/00-General/UserGroup/prg_User.TcPOU
PROGRAM prg_User
VAR
	actUser: E_userGroup:=1;
		
	ton_UserLoged: TON;
	Password: INT;
	ton_Password: TON;
	PT: BOOL;
END_VAR

ton_UserLoged(IN:=actUser<>Group1, PT:=T#10M);

IF ton_UserLoged.Q OR Password=1  THEN
	actUser:=1;
END_IF

IF Password=726 THEN
	actUser:=2;
END_IF

IF Password=345 THEN
	actUser:=3;
END_IF

IF Password=888 THEN
	actUser:=4;
END_IF


ton_Password(IN:=Password<> 0, PT:=T#1s);
IF ton_Password.Q THEN
	Password:=0;
END_IF
;

END_PROGRAM

// ---- 03 Project/23 CIP/FB_CIP_Source.TcPOU
FUNCTION_BLOCK FB_CIP_Source EXTENDS FB_SFC_Cycle IMPLEMENTS ITF_FB_SFC_Cycle
VAR_INPUT
	//eElementID			: E_Element_List;
	
	valTank_Water			: E_Pis_Name;
	valTank_R_Water			: E_Pis_Name;
	valTank_Detergent		: E_Pis_Name;
	valTank_DisInfection	: E_Pis_Name;	
	valDrain				: E_Pis_Name;
END_VAR
VAR_OUTPUT
END_VAR
VAR
	//refElement		: REFERENCE TO FB_Element;
	//refState_Long		: REFERENCE TO E_Element_State_Long;
	eReq				: E_CIP_Source;
	eProcess			: E_CIP_Source;
	eStatus				: E_CIP_Source;
	
	fbPis					: FB_Piston;
	stPis_Tank_Water		: REFERENCE TO ST_Piston;
	stPis_Tank_R_Water		: REFERENCE TO ST_Piston;
	stPis_Tank_Detergent	: REFERENCE TO ST_Piston;
	stPis_Tank_DisInfection	: REFERENCE TO ST_Piston;
	stPis_Drain				: REFERENCE TO ST_Piston;
	rt_Req_Reset: R_TRIG;
END_VAR
VAR_IN_OUT


END_VAR

act_GetReference();

act_Oper();
IF NOT Init.x THEN;
	act_Status();
END_IF

m_Request_Reset(memo:=rt_Req_Reset);//

ACTION _aClose_active:
bStepDone:=FALSE;
IF TRUE 
AND eStatus=E_CIP_Source.eClose
THEN;
	bStepDone:=TRUE;
END_IF
END_ACTION

ACTION _aClose_entry:
fbPis.m_SetByRecipe(stPis:=stPis_Tank_Water, 			req:=E_Piston_Recipe_State.Release);
fbPis.m_SetByRecipe(stPis:=stPis_Tank_R_Water, 			req:=E_Piston_Recipe_State.Release);
fbPis.m_SetByRecipe(stPis:=stPis_Tank_Detergent, 		req:=E_Piston_Recipe_State.Release);
fbPis.m_SetByRecipe(stPis:=stPis_Tank_DisInfection, 	req:=E_Piston_Recipe_State.Release);
fbPis.m_SetByRecipe(stPis:=stPis_Drain, 				req:=E_Piston_Recipe_State.Release);
END_ACTION

ACTION _aDetergent_entry:
fbPis.m_SetByRecipe(stPis:=stPis_Tank_Water, 			req:=E_Piston_Recipe_State.Release);
fbPis.m_SetByRecipe(stPis:=stPis_Tank_R_Water, 			req:=E_Piston_Recipe_State.Release);
fbPis.m_SetByRecipe(stPis:=stPis_Tank_Detergent, 		req:=E_Piston_Recipe_State.Act);
fbPis.m_SetByRecipe(stPis:=stPis_Tank_DisInfection, 	req:=E_Piston_Recipe_State.Release);
//fbPis.m_SetByRecipe(stPis:=stPis_Drain, 				req:=E_Piston_Recipe_State.Act);
END_ACTION

ACTION _aDone_entry:
eProcess:=E_CIP_Source.eNone;
eReq:=E_CIP_Source.eNone;
bRun:=FALSE;
bDone:=TRUE;
END_ACTION

ACTION _aInit_active:
SFCReset:=FALSE;
END_ACTION

ACTION _aInit_exit:
eProcess:=E_CIP_Source.eNone;
eReq:=E_CIP_Source.eNone;
END_ACTION

ACTION _aR_Water_entry:
fbPis.m_SetByRecipe(stPis:=stPis_Tank_Water, 			req:=E_Piston_Recipe_State.Release);
fbPis.m_SetByRecipe(stPis:=stPis_Tank_R_Water, 			req:=E_Piston_Recipe_State.Act);
fbPis.m_SetByRecipe(stPis:=stPis_Tank_Detergent, 		req:=E_Piston_Recipe_State.Release);
fbPis.m_SetByRecipe(stPis:=stPis_Tank_DisInfection, 	req:=E_Piston_Recipe_State.Release);
//fbPis.m_SetByRecipe(stPis:=stPis_Drain, 				req:=E_Piston_Recipe_State.Act);
END_ACTION

ACTION _aReady_active:


CASE eReq OF
	E_CIP_Source.eClose:;
			IF TRUE THEN;
				eProcess:=E_CIP_Source.eClose;
			END_IF

	E_CIP_Source.eT91_Sanitation:;
			IF TRUE THEN;
				eProcess:=E_CIP_Source.eT91_Sanitation;
			END_IF	
			
	E_CIP_Source.eT92_Detergent:;
			IF TRUE THEN;
				eProcess:=E_CIP_Source.eT92_Detergent;
			END_IF	

	E_CIP_Source.eT93_R_Water:;
			IF TRUE THEN;
				eProcess:=E_CIP_Source.eT93_R_Water;
			END_IF	
			
	E_CIP_Source.eT94_Water:;
			IF TRUE THEN;
				eProcess:=E_CIP_Source.eT94_Water;
			END_IF	

END_CASE
END_ACTION

ACTION _aReady_entry:

END_ACTION

ACTION _aReady_exit:
bRun:=TRUE;
bDone:=FALSE;
END_ACTION

ACTION _aSanitation_entry:
fbPis.m_SetByRecipe(stPis:=stPis_Tank_Water, 			req:=E_Piston_Recipe_State.Release);
fbPis.m_SetByRecipe(stPis:=stPis_Tank_R_Water, 			req:=E_Piston_Recipe_State.Release);
fbPis.m_SetByRecipe(stPis:=stPis_Tank_Detergent, 		req:=E_Piston_Recipe_State.Release);
fbPis.m_SetByRecipe(stPis:=stPis_Tank_DisInfection, 	req:=E_Piston_Recipe_State.Act);
END_ACTION

ACTION _aT91_Drain_Done_active:
bStepDone:=FALSE;
IF TRUE 
AND eStatus=E_CIP_Source.eT91_Sanitation
THEN;
	bStepDone:=TRUE;
END_IF
END_ACTION

ACTION _aT91_Drain_Done_entry:
fbPis.m_SetByRecipe(stPis:=stPis_Drain, 				req:=E_Piston_Recipe_State.Act);
END_ACTION

ACTION _aT92_Drain_Done_active:
bStepDone:=FALSE;
IF TRUE 
AND eStatus=E_CIP_Source.eT92_Detergent
THEN;
	bStepDone:=TRUE;
END_IF
END_ACTION

ACTION _aT92_Drain_Done_entry:
fbPis.m_SetByRecipe(stPis:=stPis_Drain, 				req:=E_Piston_Recipe_State.Act);
END_ACTION

ACTION _aT93_Drain_Done_active:
bStepDone:=FALSE;
IF TRUE 
AND eStatus=E_CIP_Source.eT93_R_Water
THEN;
	bStepDone:=TRUE;
END_IF
END_ACTION

ACTION _aT93_Drain_Done_entry:
fbPis.m_SetByRecipe(stPis:=stPis_Drain, 				req:=E_Piston_Recipe_State.Act);
END_ACTION

ACTION _aWater_active:
bStepDone:=FALSE;
IF TRUE 
AND eStatus=E_CIP_Source.eT94_Water
THEN;
	bStepDone:=TRUE;
END_IF
END_ACTION

ACTION _aWater_entry:
fbPis.m_SetByRecipe(stPis:=stPis_Tank_Water, 			req:=E_Piston_Recipe_State.Act);
fbPis.m_SetByRecipe(stPis:=stPis_Tank_R_Water, 			req:=E_Piston_Recipe_State.Release);
fbPis.m_SetByRecipe(stPis:=stPis_Tank_Detergent, 		req:=E_Piston_Recipe_State.Release);
fbPis.m_SetByRecipe(stPis:=stPis_Tank_DisInfection, 	req:=E_Piston_Recipe_State.Release);
fbPis.m_SetByRecipe(stPis:=stPis_Drain, 				req:=E_Piston_Recipe_State.Release);
END_ACTION

ACTION act_GetReference:
m_Set_SFCFlags_Reference();
//refElement REF= fbElement[eElementID];
//refState_Long REF= fbElement[eElementID].eState_Long;
	
stPis_Tank_Water			REF= g_Piston.stPis[valTank_Water];
stPis_Tank_R_Water			REF= g_Piston.stPis[valTank_R_Water];
stPis_Tank_Detergent		REF= g_Piston.stPis[valTank_Detergent];
stPis_Tank_DisInfection		REF= g_Piston.stPis[valTank_DisInfection];
stPis_Drain					REF= g_Piston.stPis[valDrain];
END_ACTION

ACTION act_Oper:
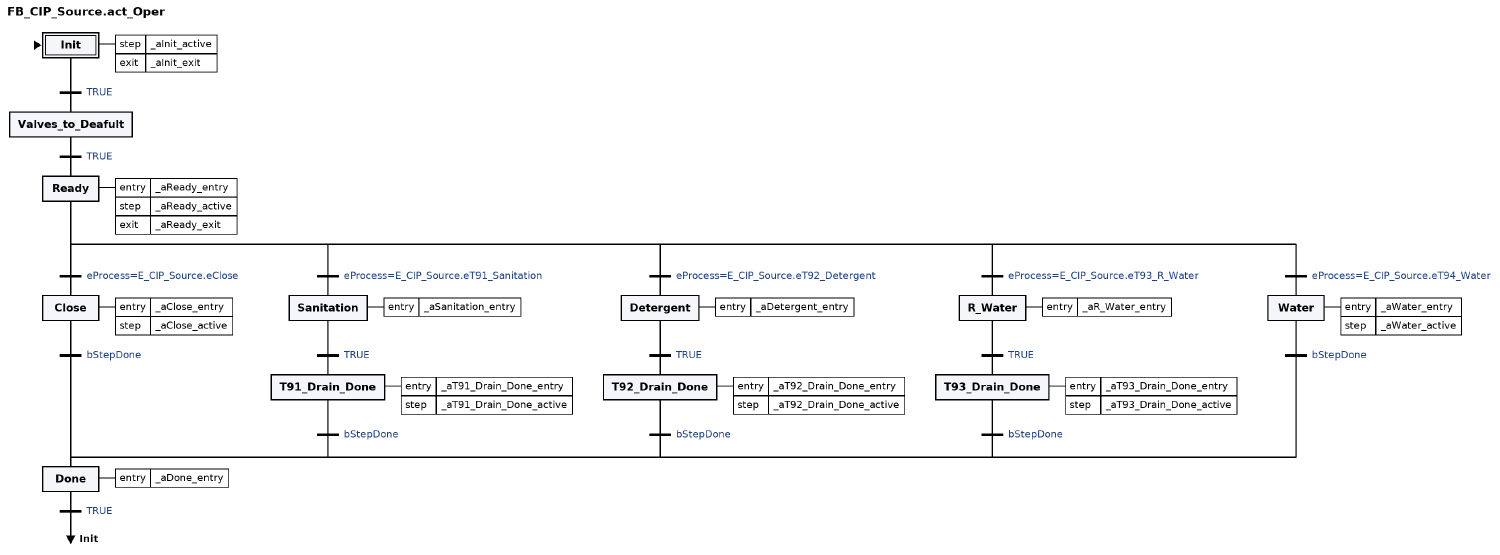
INITIAL_STEP Init:  // min time T#0.5s
    _aInit_active(N);  // step action
    _aInit_exit(P0);  // exit action
END_STEP
TRANSITION FROM Init TO Valves_to_Deafult
    := TRUE;
END_TRANSITION
STEP Valves_to_Deafult:
END_STEP
TRANSITION FROM Valves_to_Deafult TO Ready
    := TRUE;
END_TRANSITION
STEP Ready:
    _aReady_entry(P1);  // entry action
    _aReady_active(N);  // step action
    _aReady_exit(P0);  // exit action
END_STEP
TRANSITION FROM Ready TO Close
    := eProcess=E_CIP_Source.eClose;
END_TRANSITION
STEP Close:
    _aClose_entry(P1);  // entry action
    _aClose_active(N);  // step action
END_STEP
TRANSITION FROM Close TO Done
    := bStepDone;
END_TRANSITION
TRANSITION FROM Ready TO Sanitation
    := eProcess=E_CIP_Source.eT91_Sanitation;
END_TRANSITION
STEP Sanitation:  // min time T#7s
    _aSanitation_entry(P1);  // entry action
END_STEP
TRANSITION FROM Sanitation TO T91_Drain_Done
    := TRUE;
END_TRANSITION
STEP T91_Drain_Done:
    _aT91_Drain_Done_entry(P1);  // entry action
    _aT91_Drain_Done_active(N);  // step action
END_STEP
TRANSITION FROM T91_Drain_Done TO Done
    := bStepDone;
END_TRANSITION
TRANSITION FROM Ready TO Detergent
    := eProcess=E_CIP_Source.eT92_Detergent;
END_TRANSITION
STEP Detergent:  // min time T#6s
    _aDetergent_entry(P1);  // entry action
END_STEP
TRANSITION FROM Detergent TO T92_Drain_Done
    := TRUE;
END_TRANSITION
STEP T92_Drain_Done:
    _aT92_Drain_Done_entry(P1);  // entry action
    _aT92_Drain_Done_active(N);  // step action
END_STEP
TRANSITION FROM T92_Drain_Done TO Done
    := bStepDone;
END_TRANSITION
TRANSITION FROM Ready TO R_Water
    := eProcess=E_CIP_Source.eT93_R_Water;
END_TRANSITION
STEP R_Water:  // min time T#5s
    _aR_Water_entry(P1);  // entry action
END_STEP
TRANSITION FROM R_Water TO T93_Drain_Done
    := TRUE;
END_TRANSITION
STEP T93_Drain_Done:
    _aT93_Drain_Done_entry(P1);  // entry action
    _aT93_Drain_Done_active(N);  // step action
END_STEP
TRANSITION FROM T93_Drain_Done TO Done
    := bStepDone;
END_TRANSITION
TRANSITION FROM Ready TO Water
    := eProcess=E_CIP_Source.eT94_Water;
END_TRANSITION
STEP Water:
    _aWater_entry(P1);  // entry action
    _aWater_active(N);  // step action
END_STEP
TRANSITION FROM Water TO Done
    := bStepDone;
END_TRANSITION
STEP Done:  // min time T#0.2s
    _aDone_entry(P1);  // entry action
END_STEP
TRANSITION FROM Done TO Init
    := TRUE;
END_TRANSITION
// branch label Branch1_act_Oper
END_ACTION

ACTION act_Status:
IF bReady AND bDone OR TRUE THEN;
	IF TRUE 
	AND fbPis.m_CheckByRecipe(stPis:=stPis_Tank_Water, 			req:=E_Piston_Recipe_State.Release)
	AND fbPis.m_CheckByRecipe(stPis:=stPis_Tank_R_Water, 		req:=E_Piston_Recipe_State.Release)
	AND fbPis.m_CheckByRecipe(stPis:=stPis_Tank_Detergent, 		req:=E_Piston_Recipe_State.Release)
	AND fbPis.m_CheckByRecipe(stPis:=stPis_Tank_DisInfection, 	req:=E_Piston_Recipe_State.Release)
	AND fbPis.m_CheckByRecipe(stPis:=stPis_Drain, 				req:=E_Piston_Recipe_State.Release)
	THEN;
		eStatus:=E_CIP_Source.eClose;
	
	ELSIF TRUE 
	AND fbPis.m_CheckByRecipe(stPis:=stPis_Tank_Water, 			req:=E_Piston_Recipe_State.Act)
	AND fbPis.m_CheckByRecipe(stPis:=stPis_Tank_R_Water, 		req:=E_Piston_Recipe_State.Release)
	AND fbPis.m_CheckByRecipe(stPis:=stPis_Tank_Detergent, 		req:=E_Piston_Recipe_State.Release)
	AND fbPis.m_CheckByRecipe(stPis:=stPis_Tank_DisInfection, 	req:=E_Piston_Recipe_State.Release)
	AND fbPis.m_CheckByRecipe(stPis:=stPis_Drain, 				req:=E_Piston_Recipe_State.Release)
	THEN;
		eStatus:=E_CIP_Source.eT94_Water;
		
	ELSIF TRUE 
	AND fbPis.m_CheckByRecipe(stPis:=stPis_Tank_Water, 			req:=E_Piston_Recipe_State.Release)
	AND fbPis.m_CheckByRecipe(stPis:=stPis_Tank_R_Water, 		req:=E_Piston_Recipe_State.Act)
	AND fbPis.m_CheckByRecipe(stPis:=stPis_Tank_Detergent, 		req:=E_Piston_Recipe_State.Release)
	AND fbPis.m_CheckByRecipe(stPis:=stPis_Tank_DisInfection, 	req:=E_Piston_Recipe_State.Release)
	AND fbPis.m_CheckByRecipe(stPis:=stPis_Drain, 				req:=E_Piston_Recipe_State.Act)
	THEN;
		eStatus:=E_CIP_Source.eT93_R_Water;
		
	ELSIF TRUE 	
	AND fbPis.m_CheckByRecipe(stPis:=stPis_Tank_Water, 			req:=E_Piston_Recipe_State.Release)
	AND fbPis.m_CheckByRecipe(stPis:=stPis_Tank_R_Water, 		req:=E_Piston_Recipe_State.Release)
	AND fbPis.m_CheckByRecipe(stPis:=stPis_Tank_Detergent, 		req:=E_Piston_Recipe_State.Act)
	AND fbPis.m_CheckByRecipe(stPis:=stPis_Tank_DisInfection, 	req:=E_Piston_Recipe_State.Release)
	AND fbPis.m_CheckByRecipe(stPis:=stPis_Drain, 				req:=E_Piston_Recipe_State.Act)
	THEN;
		eStatus:=E_CIP_Source.eT92_Detergent;
		
